(* IEC 61131-3 sources: daoli-st-library/DL_Process (part 69) *)

(* ---- FB_DL_PressFitStation.st ---- *)
(*==============================================================================
 * 组件名称 (Component)  : FB_DL_PressFitStation
 * 所属子库 (Sublibrary) : DL_Process
 * 当前版本 (Version)    : 1.0.0
 * 组件分类 (Category)   : 功能块（FUNCTION_BLOCK）· 工站模板 · 伺服精密压装
 * 兼容性 (Platform)     : CODESYS 3.5 / TwinCAT 3 / 汇川 InoProShop / Machine Expert；
 *                         仅依赖标准库（TON / R_TRIG / ABS / LIMIT / MAX / MIN），
 *                         位移与压力均为引脚注入的工程量，块内零硬件与零轴库细节
 * 功能描述 (Function)   : 伺服精密压装工站八态（待机 / 接近 / 压入 / 保压 / 回退 /
 *                         判定 / 完成 / 故障）；压入过程逐点做位移-压力包络窗口校验
 *                         （上下限按位移节点线性插值），提取接触点 / 屈服点 / 峰值点
 *                         / 终点四特征点，一个循环给出合格结论与 NG 原因位
 * 与既有件边界 (Scope)  : 轴级力矩限幅与到位判定属运动层力矩限幅件（只出「达限 /
 *                         到位」两个布尔）；本块做工站级工艺判定（包络 + 曲线特征 +
 *                         多原因归并 + 结果结构），分层不同、不可互替。通用步序基类
 *                         不套用：压装态与监控量强耦合，套基类会出现两套状态机并存
 * 状态机规模 (States)   : 八态最小子集（0 / 10 / 20 / 30 / 40 / 50 / 60 / 99），编号
 *                         留 10 间隔便于插态；不重复包装机十七态全集（那由包装机
 *                         状态机件承担），本块只做压装工序自身的可执行子集
 * 采样口径 (Sampling)   : 接近 / 压入 / 保压三段逐拍采样；包络校验只在压入与保压段
 *                         执行（接近段压力天然低于下限，一并判会误报）；斜率按相邻
 *                         两拍差分，位移增量小于保护阈值时沿用上一拍，杜绝除零
 * 屈服判据 (Yield note) : 取「斜率回落至峰值斜率的指定比例」，不以压力绝对过峰为前
 *                         提。现场屈服段多为斜率软化而非压力下降（铝壳 / 塑料件尤
 *                         甚），强求过峰则单调上升曲线永远判不出；过峰另有独立标志
 * 设计要点 (Key notes)  : ① 单拍三律：bDone 每拍预清零、eFinish 唯一置位、转出拍不
 *                           再置位；合格与不合格在 eEvaluate 一次锁存，同循环闭环
 *                         ② 包络表只读：注入表一律不改写，上下限对调在块内镜像纠正
 *                         ③ 二分定位：带防死锁计数的二分查找，节点上限 32，最多五轮
 *                         ④ 非有限值防御：位移或压力非有限时当拍拒绝采样并转故障
 *                         ⑤ 回退快照：进回退态首拍取终点特征，位置最多滞后一个扫描
 * 码位表 (Error codes)  :
 *   16#0005_01C0【信息级】包络表点数超上限已钳位为 32，不置故障位
 *   16#0005_01C1【信息级】包络上下限对调已在块内镜像修复，不置故障位
 *   16#0005_02C0【故障级】非法状态兜底
 *   16#0005_02C1【故障级】包络表非法（节点数小于 2、或位移非严格单调递增）
 *   16#0005_02C2【故障级】阶段超时（接近 / 压入 / 保压 三段共用该码）
 *   16#0005_02C3【故障级】采样非有限值（当拍拒绝更新并转故障）
 * NG 原因位 (NG bits)   : bit0 上包络越界｜bit1 下包络越界｜bit2 终点未达｜bit3 接触
 *                         未建立｜bit4 保压压降超限；按位或累计，一个循环可多位置位
 * R32 写入点次序审计 :
 *   nSampleCnt   : ① 启动拍清零（eIdle）→ ② 采样块自增（唯一自增点）
 *   uNgReason    : ① 启动拍清零 → ② 上包络越界 → ③ 下包络越界 → ④ 保压压降（eDwell
 *                  转出）→ ⑤ 终点未达（回退首拍）→ ⑥ 接触未建立（eEvaluate）→ ⑦ 复
 *                  位清；全部按位或置位，同拍按 ②③④⑤ 累加，结构上不可能互相覆盖
 *   _uErrorIdInt : ① 启动拍清零 → ② 包络表非法（启动校验）→ ③ 阶段超时（三态各一处，
 *                  同拍只命中一处）→ ④ 采样非有限 → ⑤ 非法状态（ELSE）→ ⑥ 复位清
 *   _eState      : 每拍只在 CASE 分支出口单点写入；CASE 之外仅两处（中止监视、使能撤
 *                  销），且均在 CASE 之前，次序固定
 * 验收向量 (Acceptance) :
 *   V1 包络插值：节点（0 毫米 上限 0 下限 0）、（10 毫米 上限 10 下限 2），实测位移
 *      5.0 毫米压力 5.5 千牛 → 插得上限 5.0 下限 1.0，上越界 0.5 千牛 → bit0 置位、
 *      最大偏差不小于 0.5 千牛（容差 1E-6）
 *   V2 接触点插值：采样（1.0 毫米, 0.02 千牛）、（1.2 毫米, 0.06 千牛），阈值 0.05
 *      千牛 → 接触位移 1.15 毫米（误差不超过 1E-4）
 *   V3 屈服点：斜率序列 20 / 18 / 9 千牛每毫米，比例 0.5（阈值 10）→ 斜率 9 出现那
 *      一拍锁存屈服点，锁存后不再更新
 *   V4 终点未达：目标 10.0 毫米，回退前最大位移 9.4 毫米 → bit2 置位、不合格、单拍脉冲
 *   V5 保压压降：保压起点 12.0 千牛、结束 8.0 千牛、判据 0.3 千牛 → 压降 4.0 千牛超限
 *      → bit4 置位
 *   V6 非法包络：节点数 1 → 码 02C1、故障锁存、不出完成脉冲
 * 开源溯源 (Origin)     : 参考 lisp 与 PLCopen 公开手册的「命令-监视-判定」三段分层与
 *                         工艺参数域命名组织，只借分类与参数域；状态机、插值、特征点
 *                         提取、码位与引脚契约为本库独立设计，clean-room 不构成衍生
 * 红线自检 (Redline)    : R1 零全局表与外部变量引用、零物理地址记号 ✓｜R2 零占位符 ✓
 *                         R3 纯 IEC 61131-3 加标准库 ✓｜R4 非有限值 / 除零 / 容差 /
 *                         判界 ✓｜R5 声明行中英双语同行注释 ✓｜R6 八成员逐一有 CASE
 *                         标签且含 ELSE 兜底 ✓｜R7 三沿两定时器 CASE 外无条件刷新 ✓
 * 修订历史 (Revision)   :
 *   2026-11-15  v1.0.0  首版入库（Round 11 · C 泳道 · 工站四件套之一）
 *============================================================================*)

(*------------------------------------------------------------------------------
 * 枚举: E_DL_PressFitState（归属 FB_DL_PressFitStation，同文件发布）
 *   八态：每个成员在下方主状态机中均有同名 CASE 标签，缺一即致命（R31）
 *-----------------------------------------------------------------------------*)
TYPE E_DL_PressFitState :
(
    eIdle      := 0,    // 待机：等启动沿，输出全复位 / Idle, awaiting start edge
    eApproach  := 10,   // 接近：等接触建立 / Approach, awaiting contact build-up
    ePress     := 20,   // 压入：包络校验与特征点逐拍提取 / Press, envelope and features per scan
    eDwell     := 30,   // 保压：保持压力并监视压降 / Dwell, hold and watch force decay
    eRetract   := 40,   // 回退：等回退到位或中止 / Retract, waiting for home or abort
    eEvaluate  := 50,   // 判定：归并 NG 原因并锁存结论 / Evaluate, merge NG reasons and latch
    eFinish    := 60,   // 完成：本拍出完成脉冲，下拍转待机 / Finish, done pulse this scan
    eFault     := 99    // 故障锁存：仅复位沿可退 / Fault latched, only a reset edge leaves
);
END_TYPE

(*------------------------------------------------------------------------------
 * 结构体: ST_DL_PressFitEnvelope（归属 FB_DL_PressFitStation）
 *   位移-压力包络表，由工艺组态注入；位移节点须严格单调递增
 *-----------------------------------------------------------------------------*)
TYPE ST_DL_PressFitEnvelope :
STRUCT
    nPoints   : INT;                        // 有效节点数 [个]，域 2~32 [Valid knot count]
    afPos     : ARRAY[1..32] OF REAL;       // 节点位移 [毫米]，严格单调递增 [Knot position, mm]
    afUpper   : ARRAY[1..32] OF REAL;       // 节点包络上限 [千牛] [Upper envelope limit, kN]
    afLower   : ARRAY[1..32] OF REAL;       // 节点包络下限 [千牛] [Lower envelope limit, kN]
END_STRUCT
END_TYPE

(*------------------------------------------------------------------------------
 * 结构体: ST_DL_PressFitResult（归属 FB_DL_PressFitStation）
 *   四特征点结果，未提取到时保持 0.0，对应 NG 原因位说明缺失原因
 *-----------------------------------------------------------------------------*)
TYPE ST_DL_PressFitResult :
STRUCT
    fContactPos   : REAL;                   // 接触点位移 [毫米] [Contact position, mm]
    fContactForce : REAL;                   // 接触点压力 [千牛] [Contact force, kN]
    fYieldPos     : REAL;                   // 屈服点位移 [毫米] [Yield position, mm]
    fYieldForce   : REAL;                   // 屈服点压力 [千牛] [Yield force, kN]
    fPeakPos      : REAL;                   // 峰值点位移 [毫米] [Peak position, mm]
    fPeakForce    : REAL;                   // 峰值点压力 [千牛] [Peak force, kN]
    fEndPos       : REAL;                   // 终点位移 [毫米] [End position, mm]
    fEndForce     : REAL;                   // 终点压力 [千牛] [End force, kN]
END_STRUCT
END_TYPE

(*------------------------------------------------------------------------------
 * 结构体: ST_DL_PressFitStat（归属 FB_DL_PressFitStation）
 *   跨周期统计，由调用方持有，本块只累加，掉电保持由上层负责
 *-----------------------------------------------------------------------------*)
TYPE ST_DL_PressFitStat :
STRUCT
    nCycleCount : UDINT;                    // 累计循环数 [次] [Cycle counter]
    nOkCount    : UDINT;                    // 累计合格数 [件] [Accepted counter]
    nNgCount    : UDINT;                    // 累计不合格数 [件] [Rejected counter]
END_STRUCT
END_TYPE

FUNCTION_BLOCK FB_DL_PressFitStation
VAR_INPUT
    bEnable            : BOOL;              // 使能，FALSE 回待机并复位输出 [Enable, FALSE resets to idle]
    bStart             : BOOL;              // 启动一个压装循环，上升沿受理 [Start one cycle on rising edge]
    bAbort             : BOOL;              // 中止并立即请求回退，上升沿受理 [Abort and retract on rising edge]
    bReset             : BOOL;              // 复位故障锁存，上升沿受理 [Reset latched fault on rising edge]
    fActPos            : REAL;              // 压头实际位移 [毫米]，量程 0.0~1000.0 [Ram position, mm]
    fActForce          : REAL;              // 压力传感器实测压力 [千牛]，量程 0.0~500.0 [Measured force, kN]
    fContactForceThr   : REAL := 0.05;      // 接触判定压力阈值 [千牛]，0 表示禁用接触点提取 [Contact threshold, kN]
    fYieldSlopeRatio   : REAL := 0.50;      // 屈服判据斜率比例 [-]，域 0.05~0.99 [Yield slope ratio]
    fPeakDropForce     : REAL := 0.30;      // 峰值后压降判定量 [千牛]，0 表示不判 [Force drop after peak, kN]
    fEndPosTarget      : REAL := 10.0;      // 终点位移目标 [毫米] [Target end position, mm]
    tStageTimeout      : TIME := T#5S;      // 单段动作超时 [毫秒]，0 表示不监控 [Per-stage timeout]
    tDwell             : TIME := T#500MS;   // 保压时间 [毫秒]，0 表示跳过保压 [Dwell time]
    fForceUpperLimit   : REAL := 180.0;     // 压力硬上限 [千牛]，达限立即转保压 [Hard force limit, kN]
END_VAR
VAR_OUTPUT
    eState             : E_DL_PressFitState; // 主状态机当前态 [-]，八态之一 [Current state]
    bBusy              : BOOL;              // 循环进行中，接近至回退为真 [Cycle in progress]
    bDone              : BOOL;              // 循环结束单拍脉冲 [-] [Single-scan done pulse]
    bOk                : BOOL;              // 判定合格，保持到下次启动 [Verdict OK held until next start]
    bNg                : BOOL;              // 判定不合格，保持到下次启动 [Verdict NG held until next start]
    bError             : BOOL;              // 故障级锁存，需复位清除 [Latched fault, cleared by reset]
    uErrorId           : UDINT;             // 事件码或故障码，0 表示无 [Event or fault code, 0 = none]
    uNgReason          : WORD;              // NG 原因位，bit0~bit4 见头注释 [NG reason bits, see header]
    stResult           : ST_DL_PressFitResult; // 曲线四特征点结果 [-] [Curve feature result]
    fEnvDevMax         : REAL;              // 全程包络最大偏差 [千牛]，趋势分析用 [Max envelope deviation, kN]
    nSampleCnt         : UDINT;             // 本循环有效采样点数 [点] [Valid sample count of this cycle]
END_VAR
VAR_IN_OUT
    stEnv              : ST_DL_PressFitEnvelope; // 包络表，组态注入，块内只读 [Envelope table, read-only here]
    stStat             : ST_DL_PressFitStat;     // 跨周期统计，调用方持有 [Persistent statistics held by caller]
END_VAR
VAR
    _eState            : E_DL_PressFitState := E_DL_PressFitState.eIdle; // 内部状态寄存器 [-]，唯一真值源 [Internal state register]
    _bInit             : BOOL := FALSE;     // 首扫标志，初值 FALSE，判据 NOT _bInit [First-scan flag, R19 pattern]
    _bFaultLatch       : BOOL;              // 故障级锁存，仅复位路径清 [Fault latch, reset path only]
    _uErrorIdInt       : UDINT;             // 故障级码寄存 [Fault-level code register]
    _uInfoCode         : UDINT;             // 本拍信息级码，每拍重算 [Transient info code]
    _bEnvValid         : BOOL;              // 包络表校验通过，启动拍重算 [Envelope validated at start]
    _nEnvPts           : INT;               // 生效包络节点数 [个]，域 2~32 [Effective knot count]
    _bContactFound     : BOOL;              // 接触点已提取 [Contact point captured]
    _bYieldFound       : BOOL;              // 屈服点已提取，只锁一次 [Yield point captured once]
    _bPeakPassed       : BOOL;              // 压力已回落过峰值 [Force passed its peak]
    _bHavePrev         : BOOL;              // 存在上一点采样 [Previous sample available]
    _bRetractSnapDone  : BOOL;              // 回退入口快照已完成 [Retract snapshot already taken]
    _fPrevPos          : REAL;              // 上一点位移 [毫米] [Previous position, mm]
    _fPrevForce        : REAL;              // 上一点压力 [千牛] [Previous force, kN]
    _fStartPos         : REAL;              // 循环起点位移 [毫米] [Cycle start position, mm]
    _fSlope            : REAL;              // 当前斜率 [千牛每毫米] [Current slope, kN/mm]
    _fSlopeMax         : REAL;              // 峰值斜率 [千牛每毫米] [Peak slope, kN/mm]
    _fPeakPos          : REAL;              // 峰值点位移 [毫米] [Peak position, mm]
    _fPeakForce        : REAL;              // 峰值点压力 [千牛] [Peak force, kN]
    _fDwellStartForce  : REAL;              // 保压起点压力 [千牛] [Dwell start force, kN]
    _fContactThrEff    : REAL;              // 生效接触阈值 [千牛] [Effective contact threshold, kN]
    _fYieldRatioEff    : REAL;              // 生效屈服比例 [-] [Effective yield ratio]
    _fPeakDropEff      : REAL;              // 生效压降判据 [千牛] [Effective drop criterion, kN]
    _fEndTgtEff        : REAL;              // 生效终点目标 [毫米] [Effective end target, mm]
    _fForceLimEff      : REAL;              // 生效压力硬上限 [千牛] [Effective force limit, kN]
    _tStageEff         : TIME;              // 生效单段超时 [毫秒] [Effective stage timeout]
    _tDwellEff         : TIME;              // 生效保压时间 [毫秒] [Effective dwell time]
    _fUp               : REAL;              // 插值包络上限 [千牛] [Interpolated upper bound, kN]
    _fLo               : REAL;              // 插值包络下限 [千牛] [Interpolated lower bound, kN]
    _fSpan             : REAL;              // 插值区间跨度 [毫米] [Interpolation span, mm]
    _fRatio            : REAL;              // 插值比例 [-] [Interpolation ratio]
    _fDelta            : REAL;              // 差分中间量 [千牛或毫米] [Difference term]
    afPosUse           : ARRAY[1..32] OF REAL;  // 位移节点镜像 [毫米] [Position knot mirror, mm]
    afUpperUse         : ARRAY[1..32] OF REAL;  // 包络上限镜像 [千牛] [Upper limit mirror, kN]
    afLowerUse         : ARRAY[1..32] OF REAL;  // 包络下限镜像 [千牛] [Lower limit mirror, kN]
    nI                 : INT;               // 通用循环索引 [索引] [Loop index]
    nGuard             : INT;               // 防死锁计数 [次] [Loop guard counter]
    nLo                : INT;               // 二分下界索引 [索引] [Binary search low index]
    nHi                : INT;               // 二分上界索引 [索引] [Binary search high index]
    nMid               : INT;               // 二分中点索引 [索引] [Binary search mid index]
    bSampleFinite      : BOOL;              // 采样值有限，当拍可采 [Sample finite verdict]
    _bStageChg         : BOOL;              // 本拍发生过阶段迁移，用于断开单段计时一拍 [Stage changed this scan]
    _eStagePrev        : E_DL_PressFitState := E_DL_PressFitState.eIdle; // 上拍状态，迁移判据用 [Previous state of last scan]
    bStageTmoIn        : BOOL;              // 单段超时输入条件，先算后调 [Stage timer input]
    bDwellTmoIn        : BOOL;              // 保压计时输入条件，先算后调 [Dwell timer input]
    fbTrigStart        : R_TRIG;            // 启动沿检测 [Start edge detector]
    fbTrigAbort        : R_TRIG;            // 中止沿检测 [Abort edge detector]
    fbTrigReset        : R_TRIG;            // 复位沿检测 [Reset edge detector]
    fbTmoStage         : TON;               // 单段超时定时器 [Stage timeout timer]
    fbTmoDwell         : TON;               // 保压计时定时器 [Dwell timer]
END_VAR
VAR CONSTANT
    DL_FLOAT_EPS       : REAL := 1.0E-6;    // 浮点判等容差 [-] [Float comparison epsilon]
    DL_SLOPE_MIN_DELTA : REAL := 1.0E-4;    // 斜率计算最小位移增量 [毫米] [Min delta for slope, mm]
    DL_ENV_MAX_POINTS  : INT  := 32;        // 包络表节点数上限 [个] [Max envelope knots]
    DL_ENV_MIN_POINTS  : INT  := 2;         // 包络表节点数下限 [个] [Min envelope knots]
    DL_MAX_LOOP        : INT  := 64;        // 循环防死锁上限 [次] [Loop guard limit]
    DL_MAX_CYCLES      : UDINT := 16#FFFF_FFFE; // 统计计数饱和上限 [次] [Counter saturation limit]
    DL_RATIO_MIN       : REAL := 0.05;      // 屈服比例域下限 [-] [Yield ratio lower bound]
    DL_RATIO_MAX       : REAL := 0.99;      // 屈服比例域上限 [-] [Yield ratio upper bound]
    DL_FORCE_MAX       : REAL := 500.0;     // 压力输入域上限 [千牛] [Force domain upper bound, kN]
    DL_POS_MAX         : REAL := 1000.0;    // 位移输入域上限 [毫米] [Position domain upper bound, mm]
    DL_REAL_MAX        : REAL := 3.4E38;    // 单精度有限值判据幅值 [-] [Finite magnitude bound]
    DL_TMO_MAX         : TIME := T#180S;    // 超时参数域上限 [毫秒] [Timeout upper bound]
    DL_NG_ENV_HIGH     : WORD := 16#0001;   // NG 原因位 bit0 上包络越界 [NG bit0, upper envelope]
    DL_NG_ENV_LOW      : WORD := 16#0002;   // NG 原因位 bit1 下包络越界 [NG bit1, lower envelope]
    DL_NG_END_POS      : WORD := 16#0004;   // NG 原因位 bit2 终点未达 [NG bit2, end not reached]
    DL_NG_NO_CONTACT   : WORD := 16#0008;   // NG 原因位 bit3 接触未建立 [NG bit3, contact missing]
    DL_NG_DWELL_DROP   : WORD := 16#0010;   // NG 原因位 bit4 保压压降超限 [NG bit4, dwell decay]
    DL_INFO_PTS_CLAMP  : UDINT := 16#0005_01C0; // 01C0 包络点数越界已钳位【信息级】 [Info, knots clamped]
    DL_INFO_LIM_SWAP   : UDINT := 16#0005_01C1; // 01C1 上下限对调已修复【信息级】 [Info, limits swapped]
    DL_ERR_STATE       : UDINT := 16#0005_02C0; // 02C0 非法状态兜底【故障级】 [Fault, illegal state]
    DL_ERR_ENV         : UDINT := 16#0005_02C1; // 02C1 包络表非法【故障级】 [Fault, invalid envelope]
    DL_ERR_STAGE_TMO   : UDINT := 16#0005_02C2; // 02C2 阶段超时【故障级】 [Fault, stage timeout]
    DL_ERR_SAMPLE      : UDINT := 16#0005_02C3; // 02C3 采样非有限值【故障级】 [Fault, non-finite sample]
END_VAR
// ==== 段 1｜单拍输出预清零（R24/R25 律①：置位前先清零，任何早退路径输出确定） / Single-scan output pre-clear, mandatory before any set point
bDone      := FALSE;                        // 完成脉冲每拍先清零 [Done pulse pre-cleared]
_uInfoCode := 16#0000_0000;                 // 信息级码每拍重算 [Info code recomputed each scan]
// ==== 段 2｜工艺参数钳位（先钳位再进逻辑，杜绝分支内出现裸数值） / Parameter clamping before any logical use, no magic numbers in logic
_fContactThrEff := LIMIT(0.0, fContactForceThr, DL_FORCE_MAX);   // 接触阈值钳位 [千牛] [Contact threshold clamped]
_fYieldRatioEff := LIMIT(DL_RATIO_MIN, fYieldSlopeRatio, DL_RATIO_MAX); // 屈服比例钳位 [-] [Yield ratio clamped]
_fPeakDropEff   := LIMIT(0.0, fPeakDropForce, DL_FORCE_MAX);     // 压降判据钳位 [千牛] [Drop criterion clamped]
_fEndTgtEff     := LIMIT(0.0, fEndPosTarget, DL_POS_MAX);        // 终点目标钳位 [毫米] [End target clamped]
_fForceLimEff   := LIMIT(DL_FLOAT_EPS, fForceUpperLimit, DL_FORCE_MAX); // 硬上限钳位 [千牛] [Force limit clamped]
_tStageEff := tStageTimeout;                // 单段超时先取引脚值 [Stage timeout from pin]
IF _tStageEff > DL_TMO_MAX THEN
    _tStageEff := DL_TMO_MAX;               // 超上限钳位 [Clamped to upper bound]
ELSIF _tStageEff < T#0S THEN
    _tStageEff := T#0S;                     // 负值归零 [Negative clamped to zero]
END_IF
_tDwellEff := tDwell;                       // 保压时间先取引脚值 [Dwell time from pin]
IF _tDwellEff > DL_TMO_MAX THEN
    _tDwellEff := DL_TMO_MAX;               // 超上限钳位 [Clamped to upper bound]
ELSIF _tDwellEff < T#0S THEN
    _tDwellEff := T#0S;                     // 负值归零 [Negative clamped to zero]
END_IF
// ==== 段 3｜沿与定时器无条件刷新（R7 红线：严禁置于 IF / CASE 分支内） / Unconditional per-cycle refresh of edges and timers, outside any branch
fbTrigStart(CLK := bStart);                 // 启动沿 [Start edge]
fbTrigAbort(CLK := bAbort);                 // 中止沿 [Abort edge]
fbTrigReset(CLK := bReset);                 // 复位沿 [Reset edge]
IF ((_eState = E_DL_PressFitState.eApproach)
 OR (_eState = E_DL_PressFitState.ePress)
 OR (_eState = E_DL_PressFitState.eDwell)) AND (NOT _bStageChg) THEN
    bStageTmoIn := TRUE;                    // 动作段计时，迁移后的第一拍断输入以清零 [Timed, broken one scan after a transition]
ELSE
    bStageTmoIn := FALSE;                   // 非动作段不计时 [Timer disabled outside motion]
END_IF
fbTmoStage(IN := bStageTmoIn, PT := _tStageEff);
IF _eState = E_DL_PressFitState.eDwell THEN
    bDwellTmoIn := TRUE;                    // 仅保压段计时 [Only during dwell]
ELSE
    bDwellTmoIn := FALSE;                   // 其余段清零 [Cleared otherwise]
END_IF
fbTmoDwell(IN := bDwellTmoIn, PT := _tDwellEff);
// ==== 段 4｜首扫初始化（R19 唯一合法范式：初值 FALSE，判据 NOT，同步后置 TRUE） / First-scan initialisation with the canonical R19 pattern
IF NOT _bInit THEN
    _eState           := E_DL_PressFitState.eIdle;  // 状态回待机 [State to idle]
    _bFaultLatch      := FALSE;             // 故障锁存清零 [Fault latch cleared]
    _uErrorIdInt      := 16#0000_0000;      // 故障码清零 [Fault code cleared]
    _bEnvValid        := FALSE;             // 包络未校验 [Envelope not validated yet]
    _bStageChg        := FALSE;             // 阶段迁移标志清零 [Stage change flag cleared]
    _eStagePrev       := E_DL_PressFitState.eIdle;  // 上拍状态同步 [Previous state synced]
    _nEnvPts          := 0;                 // 节点数清零 [Knot count cleared]
    _bContactFound    := FALSE;  _bYieldFound   := FALSE;   // 接触点与屈服点未提取 [Contact and yield not captured]
    _bPeakPassed      := FALSE;  _bHavePrev     := FALSE;   // 过峰标志与采样链清零 [Peak flag and sampling chain cleared]
    _bRetractSnapDone := FALSE;             // 回退快照未做 [Retract snapshot pending]
    _fPrevPos         := 0.0;    _fPrevForce    := 0.0;     // 上一点位移与压力清零 [Previous sample cleared]
    _fStartPos        := 0.0;    _fDwellStartForce := 0.0;  // 起点与保压起点压力清零 [Start points cleared]
    _fSlope           := 0.0;    _fSlopeMax     := 0.0;     // 斜率与峰值斜率清零 [Slope and peak slope cleared]
    _fPeakPos         := 0.0;    _fPeakForce    := 0.0;     // 峰值点清零 [Peak point cleared]
    fEnvDevMax        := 0.0;    _fUp           := 0.0;     // 最大偏差与插值上限清零 [Deviation and upper bound cleared]
    _fLo              := 0.0;                               // 插值下限清零 [Lower bound cleared]
    bOk               := FALSE;  bNg            := FALSE;   // 合格与不合格结论清零 [Verdicts cleared]
    bBusy             := FALSE;  bError         := FALSE;   // 忙与故障标志清零 [Busy and error cleared]
    uErrorId          := 16#0000_0000;  uNgReason := 16#0000;  // 事件码与原因位清零 [Error id and NG bits cleared]
    nSampleCnt        := 0;                 // 采样计数清零 [Sample counter cleared]
    stResult.fContactPos   := 0.0;  stResult.fContactForce := 0.0;  // 接触点清零 [Contact point cleared]
    stResult.fYieldPos     := 0.0;  stResult.fYieldForce   := 0.0;  // 屈服点清零 [Yield point cleared]
    stResult.fPeakPos      := 0.0;  stResult.fPeakForce    := 0.0;  // 峰值点清零 [Peak point cleared]
    stResult.fEndPos       := 0.0;  stResult.fEndForce     := 0.0;  // 终点清零 [End point cleared]
    FOR nI := 1 TO DL_ENV_MAX_POINTS DO
        afPosUse[nI]   := 0.0;              // 位移镜像清零 [Position mirror cleared]
        afUpperUse[nI] := 0.0;              // 上限镜像清零 [Upper mirror cleared]
        afLowerUse[nI] := 0.0;              // 下限镜像清零 [Lower mirror cleared]
    END_FOR
    _bInit := TRUE;                         // 首扫只做一次 [Runs exactly once]
END_IF
// ==== 段 5｜启动拍包络表校验（只读校验，上下限对调在镜像里纠正，绝不改写组态） / Envelope validation at start; swaps are repaired in the mirror only
IF fbTrigStart.Q AND (_eState = E_DL_PressFitState.eIdle)
AND bEnable AND (NOT _bFaultLatch) THEN
    _bEnvValid := TRUE;                     // 先假定合法，再逐条反证 [Assume valid, then disprove]
    _nEnvPts   := stEnv.nPoints;            // 取组态节点数 [Knot count from configuration]
    IF _nEnvPts > DL_ENV_MAX_POINTS THEN
        _nEnvPts   := DL_ENV_MAX_POINTS;    // 超上限钳到 32 [Clamped to 32]
        _uInfoCode := DL_INFO_PTS_CLAMP;    // 01C0 点数越界已钳位【信息级】 [Info, knots clamped]
    END_IF
    IF _nEnvPts < DL_ENV_MIN_POINTS THEN
        _bEnvValid := FALSE;                // 少于两点无法插值 [Less than two knots is unusable]
    END_IF
    IF _bEnvValid THEN
        FOR nI := 1 TO _nEnvPts DO
            afPosUse[nI] := stEnv.afPos[nI];    // 位移镜像复制 [Copy position knot]
            IF stEnv.afUpper[nI] < stEnv.afLower[nI] THEN
                afUpperUse[nI] := stEnv.afLower[nI];   // 上限取原下限 [Upper takes old lower]
                afLowerUse[nI] := stEnv.afUpper[nI];   // 下限取原上限 [Lower takes old upper]
                _uInfoCode     := DL_INFO_LIM_SWAP;    // 01C1 上下限对调已修复【信息级】 [Info, limits swapped]
            ELSE
                afUpperUse[nI] := stEnv.afUpper[nI];  afLowerUse[nI] := stEnv.afLower[nI];  // 正常复制上下限 [Copy limits as-is]
            END_IF
        END_FOR
        FOR nI := 1 TO (_nEnvPts - 1) DO
            IF afPosUse[nI + 1] <= afPosUse[nI] THEN
                _bEnvValid := FALSE;        // 位移非严格单调，二分不可用 [Non-monotonic, binary search unsafe]
            END_IF
        END_FOR
    END_IF
    IF NOT _bEnvValid THEN
        _bFaultLatch := TRUE;               // 故障锁存 [Fault latched]
        _uErrorIdInt := DL_ERR_ENV;         // 02C1 包络表非法【故障级】 [Fault, invalid envelope]
        _eState      := E_DL_PressFitState.eFault;
    END_IF
END_IF
// ==== 段 6｜采样有限性防御与中止监视（全局，优先于状态机） / Sample finiteness defense and abort monitor, ahead of the state machine
bSampleFinite := (fActPos >= (-DL_REAL_MAX)) AND (fActPos <= DL_REAL_MAX)
             AND (fActForce >= (-DL_REAL_MAX)) AND (fActForce <= DL_REAL_MAX);
IF bEnable AND (NOT _bFaultLatch)
AND (_eState <> E_DL_PressFitState.eIdle)
AND (_eState <> E_DL_PressFitState.eFault)
AND (NOT bSampleFinite) THEN
    _bFaultLatch := TRUE;                   // 非有限值属故障级，立即锁存 [Non-finite is a fault]
    _uErrorIdInt := DL_ERR_SAMPLE;          // 02C3 采样非有限值【故障级】 [Fault, non-finite sample]
    _eState      := E_DL_PressFitState.eFault;
END_IF

IF bEnable AND (NOT _bFaultLatch) AND fbTrigAbort.Q
AND ((_eState = E_DL_PressFitState.eApproach)
  OR (_eState = E_DL_PressFitState.ePress)
  OR (_eState = E_DL_PressFitState.eDwell)) THEN
    _bHavePrev := FALSE;                    // 中止后重新起算差分 [Difference restarts after abort]
    _eState    := E_DL_PressFitState.eRetract;
END_IF
// ==== 段 7｜使能撤销（FALSE 立即回待机并撤全部动作出口，保留故障锁存） / Disable path returns to idle immediately, fault latch is preserved
IF NOT bEnable THEN
    _eState      := E_DL_PressFitState.eIdle;
    _bHavePrev   := FALSE;                  // 采样链断，防跨循环沿用 [Sampling chain broken]
    bBusy        := FALSE;                  // 忙标志撤 [Busy withdrawn]
END_IF
// ==== 段 8｜采样与特征点提取（接近 / 压入 / 保压三段逐拍执行） / Sampling and feature extraction, one sample per scan in three stages
IF bEnable AND (NOT _bFaultLatch) AND bSampleFinite
AND ((_eState = E_DL_PressFitState.eApproach)
  OR (_eState = E_DL_PressFitState.ePress)
  OR (_eState = E_DL_PressFitState.eDwell)) THEN

    IF _bHavePrev THEN
        // ---- 斜率：相邻两拍差分，位移增量过小时沿用上一拍，杜绝除零
        _fDelta := fActPos - _fPrevPos;
        IF ABS(_fDelta) >= DL_SLOPE_MIN_DELTA THEN
            _fSlope := (fActForce - _fPrevForce) / _fDelta;   // 斜率 [千牛每毫米] [Slope, kN/mm]
        END_IF
        IF _fSlope > _fSlopeMax THEN
            _fSlopeMax := _fSlope;          // 跟踪峰值斜率 [Track peak slope]
        END_IF
        // ---- 接触点：首个越过阈值的采样，用相邻两采样线性插值求精确位移
        IF (NOT _bContactFound) AND (_fContactThrEff > DL_FLOAT_EPS)
        AND (fActForce >= _fContactThrEff) THEN
            _fDelta := fActForce - _fPrevForce;
            IF ABS(_fDelta) > DL_FLOAT_EPS THEN
                stResult.fContactPos := _fPrevPos
                    + (fActPos - _fPrevPos) * (_fContactThrEff - _fPrevForce) / _fDelta;
            ELSE
                stResult.fContactPos := fActPos;   // 压力已稳定在阈值上，退化为当前点 [Degenerate to current point]
            END_IF
            stResult.fContactForce := fActForce;   // 接触点压力 [Contact force, kN]
            _bContactFound         := TRUE;        // 只锁一次 [Latched once]
        END_IF
    END_IF

    // ---- 峰值点：全程最大压力及其位移，逐拍刷新
    IF fActForce > _fPeakForce THEN
        _fPeakForce        := fActForce;    // 峰值压力 [千牛] [Peak force, kN]
        _fPeakPos          := fActPos;      // 峰值位移 [毫米] [Peak position, mm]
        stResult.fPeakForce := _fPeakForce;
        stResult.fPeakPos   := _fPeakPos;
    END_IF
    IF fActForce < (_fPeakForce - DL_FLOAT_EPS) THEN
        _bPeakPassed := TRUE;               // 已回落过峰值，趋势用 [Force has passed its peak]
    END_IF

    // ---- 屈服点：斜率回落至峰值斜率指定比例，首次成立即锁存
    IF (NOT _bYieldFound) AND _bContactFound AND (_fSlopeMax > DL_FLOAT_EPS) THEN
        IF _fSlope < (_fSlopeMax * _fYieldRatioEff) THEN
            stResult.fYieldPos   := fActPos;    // 屈服位移 [毫米] [Yield position, mm]
            stResult.fYieldForce := fActForce;  // 屈服压力 [千牛] [Yield force, kN]
            _bYieldFound         := TRUE;       // 只锁一次 [Latched once]
        END_IF
    END_IF

    nSampleCnt := nSampleCnt + 1;           // 有效采样计数 [Valid sample counter]
    _fPrevPos  := fActPos;                  // 上一点位移刷新 [Previous position refreshed]
    _fPrevForce := fActForce;               // 上一点压力刷新 [Previous force refreshed]
    _bHavePrev := TRUE;                     // 已有上一点 [Previous sample available]

    // ---- 包络窗口校验：仅压入与保压段，接近段压力天然低于下限故不判
    IF (_eState = E_DL_PressFitState.ePress) OR (_eState = E_DL_PressFitState.eDwell) THEN
        nLo    := 1;
        nHi    := _nEnvPts;
        nGuard := 0;
        WHILE ((nHi - nLo) > 1) AND (nGuard < DL_MAX_LOOP) DO
            nGuard := nGuard + 1;           // 防死锁计数 [Guard incremented]
            nMid   := (nLo + nHi) / 2;      // 整数中点 [Integer midpoint]
            IF fActPos >= afPosUse[nMid] THEN
                nLo := nMid;                // 落在右半区 [Right half]
            ELSE
                nHi := nMid;                // 落在左半区 [Left half]
            END_IF
        END_WHILE
        _fSpan := afPosUse[nHi] - afPosUse[nLo];
        IF ABS(_fSpan) > DL_SLOPE_MIN_DELTA THEN
            _fRatio := (fActPos - afPosUse[nLo]) / _fSpan;         // 区间内比例 [-] [Ratio in interval]
            _fRatio := LIMIT(0.0, _fRatio, 1.0);                   // 区间外钳位 [Clamped to 0..1]
            _fUp := afUpperUse[nLo] + _fRatio * (afUpperUse[nHi] - afUpperUse[nLo]); // 插值上限 [Interpolated upper]
            _fLo := afLowerUse[nLo] + _fRatio * (afLowerUse[nHi] - afLowerUse[nLo]); // 插值下限 [Interpolated lower]
        ELSE
            _fUp := afUpperUse[nLo];        // 退化区间取左节点上限 [Degenerate, take left knot]
            _fLo := afLowerUse[nLo];        // 退化区间取左节点下限 [Degenerate, take left knot]
        END_IF
        IF fActForce > (_fUp + DL_FLOAT_EPS) THEN
            uNgReason := uNgReason OR DL_NG_ENV_HIGH;              // bit0 上包络越界 [Upper envelope violated]
            IF (fActForce - _fUp) > fEnvDevMax THEN
                fEnvDevMax := fActForce - _fUp;                    // 累计最大偏差 [Track max deviation]
            END_IF
        END_IF
        IF fActForce < (_fLo - DL_FLOAT_EPS) THEN
            uNgReason := uNgReason OR DL_NG_ENV_LOW;               // bit1 下包络越界 [Lower envelope violated]
            IF (_fLo - fActForce) > fEnvDevMax THEN
                fEnvDevMax := _fLo - fActForce;                    // 累计最大偏差 [Track max deviation]
            END_IF
        END_IF
    END_IF
END_IF
// ==== 段 9｜主状态机（ENUM 加 CASE 加 ELSE 兜底，八成员逐一有标签） / Main state machine, every enum member has its own label
CASE _eState OF
    E_DL_PressFitState.eIdle: // 待机：等启动沿，启动拍清循环量
        IF fbTrigStart.Q AND bEnable AND (NOT _bFaultLatch) AND _bEnvValid THEN
            uNgReason    := 16#0000;  fEnvDevMax := 0.0;  nSampleCnt := 0;   // 原因位、最大偏差、采样计数清零 [Bits, deviation, count cleared]
            _bContactFound := FALSE;  _bYieldFound := FALSE;  _bPeakPassed := FALSE;  // 特征点与过峰标志复位 [Feature flags reset]
            _bHavePrev := FALSE;      _fSlope := 0.0;   _fSlopeMax := 0.0;         // 采样链、斜率、峰值斜率复位 [Chain and slope reset]
            _fPeakPos := 0.0;         _fPeakForce := 0.0;                          // 峰值点复位 [Peak reset]
            _fStartPos := fActPos;    _bRetractSnapDone := FALSE;                  // 记循环起点并复位回退快照 [Start point and snapshot reset]
            _uErrorIdInt := 16#0000_0000;  bOk := FALSE;  bNg := FALSE;            // 故障码与结论复位（启动前必无故障）[Code and verdicts reset]
            stResult.fContactPos := 0.0;  stResult.fContactForce := 0.0;           // 接触点复位 [Contact reset]
            stResult.fYieldPos   := 0.0;  stResult.fYieldForce   := 0.0;           // 屈服点复位 [Yield reset]
            stResult.fPeakPos    := 0.0;  stResult.fPeakForce    := 0.0;           // 峰值点复位 [Peak reset]
            stResult.fEndPos     := 0.0;  stResult.fEndForce     := 0.0;           // 终点复位 [End reset]
            _eState := E_DL_PressFitState.eApproach;
        END_IF
    E_DL_PressFitState.eApproach: // 接近：接触建立即转压入，阈值禁用时直通
        IF (_fContactThrEff <= DL_FLOAT_EPS) OR _bContactFound THEN
            _eState := E_DL_PressFitState.ePress;
        ELSIF fbTmoStage.Q THEN
            _bFaultLatch := TRUE;           // 阶段超时锁存 [Stage timeout latched]
            _uErrorIdInt := DL_ERR_STAGE_TMO;  // 02C2 阶段超时【故障级】 [Fault, stage timeout]
            _eState      := E_DL_PressFitState.eFault;
        END_IF
    E_DL_PressFitState.ePress: // 压入：到达终点目标或压力硬上限即转保压
        IF (fActPos >= (_fEndTgtEff - DL_FLOAT_EPS)) OR (fActForce >= _fForceLimEff) THEN
            _fDwellStartForce := fActForce; // 保压起点压力快照 [Dwell start force snapshot]
            _eState           := E_DL_PressFitState.eDwell;
        ELSIF fbTmoStage.Q THEN
            _bFaultLatch := TRUE;           // 阶段超时锁存 [Stage timeout latched]
            _uErrorIdInt := DL_ERR_STAGE_TMO;  // 02C2 阶段超时【故障级】 [Fault, stage timeout]
            _eState      := E_DL_PressFitState.eFault;
        END_IF
    E_DL_PressFitState.eDwell: // 保压：计时到即判压降并转回退，零时长直通
        IF (_tDwellEff <= T#0S) OR fbTmoDwell.Q THEN
            IF (_fPeakDropEff > DL_FLOAT_EPS)
            AND ((_fDwellStartForce - fActForce) > _fPeakDropEff) THEN
                uNgReason := uNgReason OR DL_NG_DWELL_DROP;  // bit4 保压压降超限 [Dwell decay violated]
            END_IF
            _bHavePrev := FALSE;            // 回退段不再算斜率 [Slope tracking stops]
            _eState    := E_DL_PressFitState.eRetract;
        ELSIF fbTmoStage.Q THEN
            _bFaultLatch := TRUE;           // 阶段超时锁存 [Stage timeout latched]
            _uErrorIdInt := DL_ERR_STAGE_TMO;  // 02C2 阶段超时【故障级】 [Fault, stage timeout]
            _eState      := E_DL_PressFitState.eFault;
        END_IF
    E_DL_PressFitState.eRetract: // 回退：首拍取终点特征，到位或中止即转判定
        IF NOT _bRetractSnapDone THEN
            stResult.fEndPos   := fActPos;  // 终点位移 [毫米] [End position, mm]
            stResult.fEndForce := fActForce; // 终点压力 [千牛] [End force, kN]
            IF fActPos < (_fEndTgtEff - DL_FLOAT_EPS) THEN
                uNgReason := uNgReason OR DL_NG_END_POS;  // bit2 终点未达 [End position not reached]
            END_IF
            _bRetractSnapDone := TRUE;      // 快照只做一次 [Snapshot taken once]
        END_IF
        IF fbTrigAbort.Q OR (fActPos <= (_fStartPos + DL_FLOAT_EPS)) THEN
            _eState := E_DL_PressFitState.eEvaluate;
        END_IF
    E_DL_PressFitState.eEvaluate: // 判定：归并原因并锁存结论，当拍转完成
        IF (_fContactThrEff > DL_FLOAT_EPS) AND (NOT _bContactFound) THEN
            uNgReason := uNgReason OR DL_NG_NO_CONTACT;  // bit3 接触未建立 [Contact never built up]
        END_IF
        bNg      := (uNgReason <> 16#0000); // 任一原因位即不合格 [Any reason bit means NG]
        bOk      := NOT bNg;                // 与不合格严格互斥 [Mutually exclusive with NG]
        _eState  := E_DL_PressFitState.eFinish;
    E_DL_PressFitState.eFinish: // 完成：本拍出完成脉冲并结算统计，下拍转待机
        bDone := TRUE;                      // 完成单拍，本拍唯一置位点 [Sole set point of the pulse]
        IF bNg THEN
            IF stStat.nNgCount < DL_MAX_CYCLES THEN
                stStat.nNgCount := stStat.nNgCount + 1;   // 不合格计数饱和累加 [NG counter, saturated]
            END_IF
        ELSE
            IF stStat.nOkCount < DL_MAX_CYCLES THEN
                stStat.nOkCount := stStat.nOkCount + 1;   // 合格计数饱和累加 [OK counter, saturated]
            END_IF
        END_IF
        IF stStat.nCycleCount < DL_MAX_CYCLES THEN
            stStat.nCycleCount := stStat.nCycleCount + 1; // 循环计数饱和累加 [Cycle counter, saturated]
        END_IF
        _bHavePrev := FALSE;                // 采样链断开，防跨循环 [Sampling chain broken]
        _eState    := E_DL_PressFitState.eIdle;
    E_DL_PressFitState.eFault: // 故障：等复位沿，复位后清码回待机
        IF fbTrigReset.Q THEN
            _bFaultLatch      := FALSE;     // 锁存解除 [Latch released]
            _uErrorIdInt      := 16#0000_0000; // 故障码清零 [Fault code cleared]
            uNgReason         := 16#0000;   // 原因位清零 [NG bits cleared]
            _bRetractSnapDone := FALSE;     // 快照标志复位 [Snapshot flag reset]
            _bHavePrev        := FALSE;     // 差分复位 [Difference reset]
            _eState           := E_DL_PressFitState.eIdle;
        END_IF

    ELSE // 非法枚举值兜底：回安全态并锁故障
        _bFaultLatch := TRUE;               // 兜底锁存 [Fallback latch]
        _uErrorIdInt := DL_ERR_STATE;       // 02C0 非法状态兜底【故障级】 [Fault, illegal state]
        _eState      := E_DL_PressFitState.eFault;
END_CASE
// ==== 段 10｜阶段迁移寄存器更新（单段超时的清零依据，与状态写入点分离） / Stage change register, drives the per-stage timer reset
_bStageChg  := (_eState <> _eStagePrev);     // 本拍是否发生迁移 [Transition happened this scan]
_eStagePrev := _eState;                      // 迁移寄存器同步 [Previous state synced]

// ==== 段 11｜出口派生（每拍重写，bError 只反映故障级，信息级码只进 uErrorId） / Outlets rewritten every scan, info codes never raise bError
eState := _eState;                          // 状态镜像 [State mirror]
bBusy  := (_eState = E_DL_PressFitState.eApproach)
       OR (_eState = E_DL_PressFitState.ePress)
       OR (_eState = E_DL_PressFitState.eDwell)
       OR (_eState = E_DL_PressFitState.eRetract);   // 执行中派生 [Busy derived]

bError := _bFaultLatch;                     // 故障级派生式（R21）[Fault-level derived form]
IF _bFaultLatch THEN
    uErrorId := _uErrorIdInt;               // 故障级码优先透出 [Fault code wins]
ELSE
    uErrorId := _uInfoCode;                 // 无故障时透出信息级码 [Info code otherwise]
END_IF
END_FUNCTION_BLOCK

(* ---- FB_DL_PressForceCurveExec.st ---- *)
(*==============================================================================
 * 组件名称 (Component)  : FB_DL_PressForceCurveExec
 * 所属子库 (Sublibrary) : DL_Process ｜ 版本 (Version) : 1.0.0 ｜ 2026-11-24
 * 兼容性   (Platform)   : CODESYS 3.5+ / TwinCAT 3 / 汇川 InoProShop / 施耐德 Machine Expert
 *                         仅依赖 IEC 61131-3 标准库（TON / R_TRIG / ABS / MIN / MAX / LIMIT），零厂商私有库
 * 功能描述 (Function)   : 压机多段力曲线执行：按 4 段配方（目标力 aSegForce / 升力速率 aSegRate /
 *                         保压时长 aSegHold）逐段执行，eRamp 以「速率 × dt」斜坡逼近目标力，
 *                         到力判据 = 指令已饱和到目标（|cmd − target| ≤ EPS）**且** 实际力反馈落进
 *                         容差带（容差 = max(0.5% × |目标力|, 0.1 kN)）→ eHold 保压 aSegHold[i]；
 *                         末段保压完成 → eRelease 按末段速率把力指令斜坡降到 0 → eDone 发 bCurveDone。
 *                         **dt 口径**：定周期采样节拍 tonDt（PT = 100ms 常数）生成步长
 *                         _fDtSec := TIME_TO_LREAL(DL_PFC_DT)，入口做 dt > EPS 闸（R4 防 dt ≤ 0）；
 *                         保压计时用 DINT 毫秒累加（_diHoldMs，每采样拍 +100ms），避免 TIME 加法跨型。
 *                         **bStart = FALSE 语义（R191 二选一，本件选「降级为安全值 + 置标志」）**：
 *                         力指令按段速率退回 0 并进 eIdle（压机力指令不得冻结保持）。
 * 接口     (Interface)  : 输入 bEnable / bStart / bReset（上升沿）/ aSegForce[1..4] / aSegRate[1..4] /
 *                         aSegHold[1..4] / nSegCnt / fForceFb / tSegTimeout；
 *                         输出 fForceCmd / nSegAct / tHoldElapsed / bCurveDone / eState（E_DL_PfcPhase）/
 *                         eCause（E_DL_PfcCause）/ bError / bValid / nSegCompleted。
 * 状态迁移表 (State Transition Table)：
 *   ① eIdle → eRamp：bEnable 且 bStart 且组态闸通过且无锁存；拍 N 进入 / 本拍行为：
 *      fForceCmd=0、nSegAct=1、nSegCompleted=0、_diHoldMs=0 / 拍 N+1 转出至 eRamp。
 *   ② eRamp → eHold：到力判据成立（指令饱和 + 反馈落带）；拍 N 进入 / 本拍行为：
 *      _diHoldMs 清零、fForceCmd 精确取目标 / 拍 N+1 转出至 eHold。
 *   ③ eHold → eRamp：_diHoldMs ≥ aSegHold[i] 且 i < nSegCnt；本拍行为：nSegAct+1、
 *      nSegCompleted+1、_diHoldMs 清零、信息级 eSegDone / 拍 N+1 转出（下一段）。
 *   ④ eHold → eRelease：_diHoldMs ≥ aSegHold[nSegCnt]（末段完成）；本拍行为：nSegCompleted+1、
 *      信息级 eCurveDoneCode / 拍 N+1 转出至 eRelease。
 *   ⑤ eRelease → eDone：|fForceCmd| ≤ EPS（已退到 0）；本拍行为：fForceCmd 精确置 0 /
 *      拍 N+1 转出至 eDone。
 *   ⑥ eDone → eIdle：(NOT bStart) OR bReset 上升沿（两条出口 R98）；本拍行为：bCurveDone 落 FALSE、
 *      力指令与段号清零 / 拍 N+1 转出至 eIdle。
 *   ⑦ eRamp → eFault：tonSeg.Q（单段超时未到力）锁存 eForceNotReached；本拍行为：fForceCmd 保持
 *      当前值直至段尾迁移闸（R21）后再全撤 / 拍 N+1 转出至 eFault。
 *   ⑧ 任一相 → eFault：组态闸失败（段数越域 / 速率 ≤ 0 / 目标力 < 0 / 保压越域 / 超时越域 /
 *      fForceFb 非有限），锁存首因。
 *   ⑨ eFault → eIdle：bReset 上升沿（R_TRIG 判 .Q）且 bEnable = FALSE（R19 穷举出口）；
 *      本拍行为：清锁存与成因、fForceCmd=0 / 拍 N+1 转出至 eIdle。
 *   ⑩ ELSE（非法枚举值）→ eFault，成因 eIllegalState（R6 兜底）。
 * 边界     (Boundary)   : ① tonDt / tonSeg / R_TRIG 全在 CASE 外无条件调用（R7）；两者 IN 均含
 *                            NOT .Q 自复位项（R188）；tonSeg 另含「(NOT _bSegReset)」断流项 ——
 *                            换段（含首段起始）当拍置 _bSegNew，次拍 _bSegReset 为真使 IN 断流，
 *                            ET 归零后再起计，故单段超时按段独立（结构性无需外部沿清零）。
 *                         ② 斜坡双向：目标高于当前则升、低于当前则降（段间降力不越界），
 *                            三步比较全用大小判据，无浮点等值比较（R4）。
 *                         ③ 到力容差为「相对 0.5% 与绝对 0.1 kN 取大」，浮点比较一律容差式。
 *                         ④ 组态域闸：nSegCnt ∈ [1,4]（越域直接故障并钳位供下标安全）；
 *                            参与执行的段（1..nSegCnt）逐段校验速率 > 0、目标力 ≥ 0、保压 ≤ 1h；
 *                            全部 4 段做非有限拒收（未参与段不判量程域，见分工声明）。
 *                         ⑤ 无除法，故无除零；无浮点等值比较；力指令出口恒为饱和值。
 *                         ⑥ 零全局耦合（无 GVL / VAR_EXTERNAL / %I / %Q，R1 / R2）。
 * 码表     (Codes)      : 本件不占用全局数字码位（R297 零码位范式）；出口为 BOOL + ENUM，
 *                         enum E_DL_PfcPhase / E_DL_PfcCause 归属本文件（全库唯一属主，R264）。
 *                         信息级（0..9）永不置 bError；故障级（10 起）赋值处与 _bFaultLatch 三行
 *                         成对（R45），锁存回放至 bReset 沿（FB33-1）。
 * 分工声明 (Scope)      : 压机液压比例阀闭环 / 伺服压力闭环归运动控制件；模具保护与吨位监视归
 *                         FB_DL_PressTonnageGuard 类件；本件只做**多段力配方开环斜坡 + 到力判定 +
 *                         保压计时**，不做力闭环 PID，也不做安全回路（安全由 PRG_IoMapping 双切断）。
 * 归属     (Ownership)  : E_DL_PfcPhase / E_DL_PfcCause 归属本文件（全库唯一定义，R264）。
 * 红线自检 (Redline)    : R1 ✓ 零 GVL ｜ R2 ✓ 零 %I/%Q ｜ R3 ✓ 纯 IEC ｜ R4 ✓ dt 闸 + 容差比较 +
 *                         非有限双判 + 无除法 ｜ R5 ✓ 逐行同行双语注释 ｜ R6 ✓ 六态 ENUM + CASE +
 *                         ELSE ｜ R7 ✓ 全部 TON/R_TRIG 在 CASE 外 ｜ R8/R9 N/A（无 METHOD）
 *                         R10 ✓ 无构造式转换 ｜ R14 ✓ 无 PROPERTY ｜ R15 ✓ 无保留字撞名
 *                         R17 ✓ 定长 ARRAY[1..4] ｜ R18 ✓ bReset 用 R_TRIG 判 .Q ｜ R19 ✓ eFault
 *                         出口 = bReset 沿 + 撤使能 ｜ R20 ✓ 到力等待相带 tSegTimeout 超时兜底
 *                         R21 ✓ 锁存与迁相分离。
 * 修订历史 (Revision)   : 2026-11-24  v1.0.0  R79-B 首版
 * 验收向量 (Acceptance) :
 *   V1 nSegCnt=2、段1 = (50 kN, 10 kN/s, T#2S)、段2 = (80 kN, 5 kN/s, T#1S)、tSegTimeout=T#30S、
 *      fForceFb 跟随 fForceCmd：eRamp 约 5s 到 50 kN → eHold（tHoldElapsed 递增到 2s）→ 段2：
 *      约 6s 到 80 kN → eHold 1s → eRelease → eDone，bCurveDone=TRUE、nSegCompleted=2。
 *   V2 nSegCnt=0（越域）→ eState=eFault、eCause=eBadConfig、bError=TRUE、fForceCmd=0；
 *      bReset 上升沿且 bEnable=FALSE → 回 eIdle、bError=FALSE。
 *   V3 aSegRate[1]=0.0（速率非正）→ eState=eFault、eCause=eBadConfig。
 *   V4 aSegForce[1]=50.0、tSegTimeout=T#5S、fForceFb 恒为 0（力建不起来）→ 5s 后
 *      eState=eFault、eCause=eForceNotReached、bError=TRUE、fForceCmd=0（故障相全撤）。
 *   V5 fForceFb = NaN → eState=eFault、eCause=eNonFinite（非有限拒收，非量程判据）。
 *   V6 eRamp 中 bStart 落 FALSE → fForceCmd 回 0、eState=eIdle、nSegAct=0（安全降级）。
 *============================================================================*)

(*-----------------------------------------------------------------------------
 * 枚举: E_DL_PfcPhase（压机力曲线相位；eFault 为安全相，仅 bReset 沿迁出）
 *----------------------------------------------------------------------------*)
TYPE E_DL_PfcPhase :
(
    eIdle    := 0,    // 空闲：力指令 0，段号清零 / Idle: force command zero, segment cleared
    eRamp    := 10,   // 斜坡相：按段速率逼近目标力 / Ramp: approach the target at the segment rate
    eHold    := 20,   // 保压相：力保持目标值并计时 / Hold: keep the target force and time it
    eRelease := 30,   // 卸力相：力指令斜坡降到 0 / Release: ramp the force command down to zero
    eDone    := 40,   // 完成相：bCurveDone 电平为 TRUE / Done: bCurveDone held high
    eFault   := 90    // 故障安全相：锁存成因，力指令回 0 / Fault safe phase: latched cause, force command zeroed
);
END_TYPE

(*-----------------------------------------------------------------------------
 * 枚举: E_DL_PfcCause（成因码；信息级 = 0..9，故障级 = 10 起）
 *----------------------------------------------------------------------------*)
TYPE E_DL_PfcCause :
(
    eNone            := 0,   // 信息级：无事件 / Info: no event
    eSegDone         := 1,   // 信息级：一段保压完成 / Info: one segment hold completed
    eCurveDoneCode   := 2,   // 信息级：曲线保压全部完成 / Info: all segment holds completed
    eReleasing       := 3,   // 信息级：进入卸力相 / Info: entering the release phase
    eBadConfig       := 10,  // 故障级：段数 / 速率 / 目标力 / 保压 / 超时越域 / Fault: segment, rate, force, hold or timeout out of domain
    eNonFinite       := 11,  // 故障级：入参非有限 / Fault: non-finite input
    eForceNotReached := 12,  // 故障级：单段超时未到力 / Fault: force not reached within the segment timeout
    eIllegalState    := 13   // 故障级：非法状态枚举值 / Fault: illegal state enum value
);
END_TYPE

FUNCTION_BLOCK FB_DL_PressForceCurveExec
VAR_INPUT
    bEnable     : BOOL := FALSE;                        // 使能：FALSE 力指令回 0 并回 eIdle / Enable, FALSE zeroes the force and returns to idle
    bStart      : BOOL := FALSE;                        // 启动（电平）：FALSE 曲线中止，力指返回 0 / Start level, FALSE aborts and ramps the force back
    bReset      : BOOL := FALSE;                        // 复位（上升沿，需同时 bEnable=FALSE）/ Reset rising edge, requires bEnable FALSE
    aSegForce   : ARRAY[1..4] OF LREAL;                 // 各段目标力（域 ≥ 0）[kN] / Per-segment target force, domain >= 0
    aSegRate    : ARRAY[1..4] OF LREAL;                 // 各段升力速率（域 > 0）[kN/s] / Per-segment force rate, domain > 0
    aSegHold    : ARRAY[1..4] OF TIME;                  // 各段保压时长（域 0..1h）[s] / Per-segment hold time, domain 0..1h
    nSegCnt     : INT := 1;                             // 实际执行段数，有效域 1..4 [段] / Effective segment count, valid domain 1..4
    fForceFb    : LREAL := 0.0;                         // 实际力反馈（来自压力/力传感器）[kN] / Actual force feedback
    tSegTimeout : TIME := T#30S;                        // 单段到力超时，域 100ms..1h [s] / Per-segment force-reach timeout
END_VAR
VAR_OUTPUT
    fForceCmd      : LREAL := 0.0;                      // 力指令出口（斜坡饱和值）[kN] / Force command outlet, saturated ramp value
    nSegAct        : INT := 0;                          // 当前段号（1 起，0 = 未开始）[段] / Current segment number, 0 means not started
    tHoldElapsed   : TIME := T#0S;                      // 当前段保压已用时长 [s] / Elapsed hold time of the current segment
    bCurveDone     : BOOL;                              // 曲线完成（电平，保持至 bStart 落或复位）[-] / Curve done, level held until start falls
    eState         : E_DL_PfcPhase;                     // 状态出口（段尾单点映射）[-] / State outlet mapped at the tail
    eCause         : E_DL_PfcCause;                     // 成因码出口（故障期锁存回放）[-] / Cause code outlet
    bError         : BOOL;                              // 故障锁存标志 [-] / Fault latch flag
    bValid         : BOOL;                              // 曲线有效回执（斜坡/保压相且无锁存）[-] / Curve validity receipt
    nSegCompleted  : INT := 0;                          // 已完成段数 [段] / Number of completed segments
END_VAR
VAR
    _eState       : E_DL_PfcPhase := E_DL_PfcPhase.eIdle;   // 内部相位（CASE 唯一写入目标）[-] / Internal phase
    _bFaultLatch  : BOOL := FALSE;                          // 故障锁存位（仅 bReset 沿清除）[-] / Fault latch bit
    _eCauseLatch  : E_DL_PfcCause := E_DL_PfcCause.eNone;    // 锁存成因码（FB33-1 锁存回放）[-] / Latched cause code
    _eCauseTmp    : E_DL_PfcCause := E_DL_PfcCause.eNone;    // 本拍首因中间量（段 6 组态闸用）[-] / First cause of this scan
    _bCfgOk       : BOOL := TRUE;                           // 组态与入参闸通过标志 [-] / Configuration gate flag
    _bResetPulse  : BOOL := FALSE;                          // bReset 上升沿快照（R18）[-] / bReset rising-edge snapshot
    _nSegClamp    : INT := 1;                               // 段数钳位值 1..4（下标安全）[段] / Clamped segment count for safe indexing
    _bSegNew      : BOOL := FALSE;                          // 本拍进入新段标志（CASE 内置位，次拍令单段超时 ET 自清）[-] / New-segment flag set inside CASE
    _bSegReset    : BOOL := FALSE;                          // 新段标志快照（段 1 取上一拍值，供 tonSeg 的 IN 断流）[-] / New-segment snapshot latching the last-scan value
    _nIdx         : INT := 1;                               // 遍历下标（FOR 专用）[段] / Loop index for FOR statements
    _diHoldMs     : DINT := 0;                              // 保压毫秒累加（DINT 防跨型溢出）[ms] / Accumulated hold milliseconds
    _fDtSec       : LREAL := 0.0;                           // 采样步长 [s] / Sampling step in seconds
    _bDtOk        : BOOL := FALSE;                          // 步长有效性（dt > EPS）[-] / Sampling step validity
    _fStep         : LREAL := 0.0;                          // 本拍斜坡增量 [kN] / Ramp increment of this scan
    _fTol         : LREAL := 0.0;                           // 到力容差 = max(0.5%×|目标|, 0.1) [kN] / Force-reach tolerance
    _bCmdAtTarget : BOOL := FALSE;                          // 指令已饱和到目标标志 [-] / Command saturated at the target
    _bFbInTol     : BOOL := FALSE;                          // 反馈落进容差带标志 [-] / Feedback inside the tolerance band
    rtReset       : R_TRIG;                                 // bReset 边沿实例（段 4 无条件调用，R18）/ bReset edge instance called unconditionally
    tonDt         : TON;                                    // 定周期采样节拍（段 4 无条件调用）/ Fixed-period sampling tick
    tonSeg        : TON;                                    // 单段到力超时（段 4 无条件调用）/ Per-segment force-reach timeout
END_VAR
VAR CONSTANT
    DL_PFC_ZERO      : LREAL := 0.0;             // 浮点零基准 [-] / Float zero base
    DL_PFC_EPS       : LREAL := 1.0E-6;          // 浮点同值/正步长容差（力指令饱和判）[-] / Float equality and positive-step tolerance
    DL_PFC_TOL_PCT   : LREAL := 0.005;           // 到力相对容差 0.5% [-] / Relative force tolerance of 0.5 percent
    DL_PFC_TOL_ABS   : LREAL := 0.1;             // 到力绝对容差 [kN] / Absolute force tolerance
    DL_PFC_SEG_MAX   : INT := 4;                 // 段数上限（数组定长）[段] / Upper bound of segments, fixed array size
    DL_PFC_ONE       : INT := 1;                 // 段号起始值 [段] / Segment numbering start
    DL_PFC_DT        : TIME := T#100MS;          // 采样节拍（斜坡步长来源）[s] / Sampling tick, the ramp step source
    DL_PFC_DT_MS     : DINT := 100;              // 采样节拍毫秒数（保压累加步长）[ms] / Sampling tick in milliseconds
    DL_PFC_T_MIN     : TIME := T#100MS;          // 超时参数下限 [s] / Lower bound of the timeout parameter
    DL_PFC_T_MAX     : TIME := T#1H;             // 超时与保压参数上限 [s] / Upper bound of timeout and hold time
    DL_PFC_MS_ZERO   : DINT := 0;                // 毫秒零基准 [-] / Millisecond zero base
END_VAR

(* —— 段 1：单拍与电平出口预置（不清锁存 / 力指令 / 段号状态，FB32-1） —— *)
bCurveDone := FALSE;                                   // 曲线完成电平每拍预清（仅 eDone 相重新置位）/ Curve-done level preset, re-armed only in eDone
_bCfgOk    := TRUE;                                    // 组态闸标志复位 / Configuration flag reset
_eCauseTmp := E_DL_PfcCause.eNone;                      // 当拍首因复位 / Scan cause reset
_bSegReset := _bSegNew;                                // 取上一拍的新段标志（本拍令 tonSeg 的 IN 断流，R188）/ Take the last-scan new-segment flag
_bSegNew   := FALSE;                                   // 新段标志每拍预清（仅换段相内置位）/ Preset the new-segment flag, set only on a segment change

(* —— 段 2：段数钳位与采样步长（标准转换，R10） —— *)
_nSegClamp := LIMIT(DL_PFC_ONE, nSegCnt, DL_PFC_SEG_MAX);            // 段数钳位 1..4 / Clamp the segment count
_fDtSec    := TIME_TO_LREAL(DL_PFC_DT);                              // 节拍换算为秒 / Sampling tick to seconds
IF _fDtSec > DL_PFC_EPS THEN
    _bDtOk := TRUE;                                                  // 步长为正：允许斜坡积分 / Positive step: ramp integration allowed
ELSE
    _bDtOk := FALSE;                                                 // 步长非正：拒绝积分（R4）/ Non-positive step: integration refused
END_IF

(* —— 段 3：全部 4 段非有限拒收（未参与段也拒 NaN / Inf，避免污染后续组态）/ —— *)
FOR _nIdx := 1 TO DL_PFC_SEG_MAX DO
    IF (aSegForce[_nIdx] <> aSegForce[_nIdx]) OR ((aSegForce[_nIdx] - aSegForce[_nIdx]) <> DL_PFC_ZERO) THEN
        _bCfgOk    := FALSE;                            // 目标力非有限 / Target force is not finite
        _eCauseTmp := E_DL_PfcCause.eNonFinite;         // 故障级：非有限入参 / Fault: non-finite input
    END_IF
    IF (aSegRate[_nIdx] <> aSegRate[_nIdx]) OR ((aSegRate[_nIdx] - aSegRate[_nIdx]) <> DL_PFC_ZERO) THEN
        _bCfgOk    := FALSE;                            // 速率非有限 / Rate is not finite
        _eCauseTmp := E_DL_PfcCause.eNonFinite;         // 故障级：非有限入参 / Fault: non-finite input
    END_IF
END_FOR
IF (fForceFb <> fForceFb) OR ((fForceFb - fForceFb) <> DL_PFC_ZERO) THEN
    _bCfgOk    := FALSE;                                // 力反馈非有限 / Force feedback is not finite
    _eCauseTmp := E_DL_PfcCause.eNonFinite;             // 故障级：非有限入参 / Fault: non-finite input
END_IF

(* —— 段 4：组态量程域闸（仅参与执行的 1..nSegCnt 段，逐段校验） —— *)
IF _bCfgOk THEN
    IF (nSegCnt < DL_PFC_ONE) OR (nSegCnt > DL_PFC_SEG_MAX) THEN
        _bCfgOk    := FALSE;                            // 段数越域 / Segment count out of domain
        _eCauseTmp := E_DL_PfcCause.eBadConfig;         // 故障级：组态非法 / Fault: bad configuration
    ELSIF (tSegTimeout < DL_PFC_T_MIN) OR (tSegTimeout > DL_PFC_T_MAX) THEN
        _bCfgOk    := FALSE;                            // 单段超时越域 / Segment timeout out of domain
        _eCauseTmp := E_DL_PfcCause.eBadConfig;         // 故障级：组态非法 / Fault: bad configuration
    ELSE
        FOR _nIdx := 1 TO _nSegClamp DO
            IF aSegRate[_nIdx] <= DL_PFC_ZERO THEN
                _bCfgOk    := FALSE;                    // 速率非正，无法斜坡 / Non-positive rate, ramp impossible
                _eCauseTmp := E_DL_PfcCause.eBadConfig; // 故障级：组态非法 / Fault: bad configuration
            END_IF
            IF aSegForce[_nIdx] < DL_PFC_ZERO THEN
                _bCfgOk    := FALSE;                    // 目标力为负 / Negative target force
                _eCauseTmp := E_DL_PfcCause.eBadConfig; // 故障级：组态非法 / Fault: bad configuration
            END_IF
            IF aSegHold[_nIdx] > DL_PFC_T_MAX THEN
                _bCfgOk    := FALSE;                    // 保压时长越上限 / Hold time above the upper bound
                _eCauseTmp := E_DL_PfcCause.eBadConfig; // 故障级：组态非法 / Fault: bad configuration
            END_IF
        END_FOR
    END_IF
END_IF

(* —— 段 5：边沿与定时器（CASE 外无条件调用，R7；IN 均含 NOT .Q 自复位，R188） —— *)
rtReset(CLK := bReset);                                // bReset 边沿无条件刷新（R18）/ bReset edge refreshed unconditionally
_bResetPulse := rtReset.Q;                             // 边沿快照 / Edge snapshot
tonDt(IN := ((_eState = E_DL_PfcPhase.eRamp) OR (_eState = E_DL_PfcPhase.eHold)
             OR (_eState = E_DL_PfcPhase.eRelease))
            AND (NOT tonDt.Q) AND (NOT _bFaultLatch),
      PT := DL_PFC_DT);                                // 执行相定周期采样节拍 / Fixed-period tick in the execution phases
tonSeg(IN := (_eState = E_DL_PfcPhase.eRamp) AND (NOT _bSegReset)
              AND (NOT tonSeg.Q) AND (NOT _bFaultLatch),
        PT := tSegTimeout);                            // 单段超时：换段次拍 IN 断流使 ET 自清（R188）

(* —— 段 6：状态机主体（唯一相位写入点；故障只置锁存，迁相由段 8 统一执行） —— *)
CASE _eState OF
    E_DL_PfcPhase.eIdle :
        fForceCmd     := DL_PFC_ZERO;                  // 空闲：力指令归零 / Idle: force command zeroed
        nSegAct       := 0;                            // 空闲：段号清零 / Idle: segment cleared
        nSegCompleted := 0;                            // 空闲：完成段数清零 / Idle: completed segments cleared
        _diHoldMs     := DL_PFC_MS_ZERO;               // 空闲：保压累计清零 / Idle: hold accumulator cleared
        IF bEnable AND bStart AND _bCfgOk AND (NOT _bFaultLatch) THEN
            fForceCmd  := DL_PFC_ZERO;                 // 迁移①：起点力为零 / Start from zero force
            nSegAct    := DL_PFC_ONE;                  // 从第 1 段开始 / Begin at segment one
            _diHoldMs  := DL_PFC_MS_ZERO;              // 保压累计清零 / Hold accumulator cleared
            _bSegNew   := TRUE;                        // 首段起始：次拍令单段超时 ET 自清 / First segment: reset the timeout on the next scan
            eCause     := E_DL_PfcCause.eNone;         // 信息级：无事件 / Info: no event
            _eState    := E_DL_PfcPhase.eRamp;         // 进入斜坡相 / Move to ramp
        END_IF

    E_DL_PfcPhase.eRamp :
        IF (NOT bEnable) OR (NOT bStart) THEN
            fForceCmd := DL_PFC_ZERO;                  // 失能：力指令回 0（安全降级）/ Disabled: force zeroed for safety
            nSegAct   := 0;                            // 段号清零 / Segment cleared
            eCause    := E_DL_PfcCause.eNone;          // 信息级：无事件 / Info: no event
            _eState   := E_DL_PfcPhase.eIdle;          // 回空闲相 / Back to idle
        ELSE
            (* 斜坡：按段速率把力指令推向目标（双向） *)
            IF tonDt.Q AND _bDtOk THEN
                _fStep := aSegRate[nSegAct] * _fDtSec; // 本拍增量 = 速率 × dt [kN]
                IF fForceCmd < aSegForce[nSegAct] THEN
                    fForceCmd := MIN(fForceCmd + _fStep, aSegForce[nSegAct]);   // 升力且不越过目标 / Ramp up without overshoot
                ELSIF fForceCmd > aSegForce[nSegAct] THEN
                    fForceCmd := MAX(fForceCmd - _fStep, aSegForce[nSegAct]);   // 降力且不越过目标 / Ramp down without overshoot
                END_IF
            END_IF
            (* 到力判据：容差 = max(0.5%×|目标|, 0.1 kN)，浮点比较一律容差式（R4） *)
            _fTol := MAX(ABS(aSegForce[nSegAct]) * DL_PFC_TOL_PCT, DL_PFC_TOL_ABS);
            _bCmdAtTarget := ABS(fForceCmd - aSegForce[nSegAct]) <= DL_PFC_EPS;   // 指令已饱和到目标
            _bFbInTol     := ABS(fForceFb - aSegForce[nSegAct]) <= _fTol;         // 反馈落进容差带
            IF _bCmdAtTarget AND _bFbInTol THEN
                fForceCmd := aSegForce[nSegAct];       // 迁移②：到力，指令精确取目标 / Reached: command set exactly
                _diHoldMs := DL_PFC_MS_ZERO;           // 保压累计清零 / Hold accumulator cleared
                eCause    := E_DL_PfcCause.eNone;      // 信息级：无事件 / Info: no event
                _eState   := E_DL_PfcPhase.eHold;      // 进入保压相 / Move to hold
            ELSIF tonSeg.Q THEN
                IF NOT _bFaultLatch THEN
                    _eCauseLatch := E_DL_PfcCause.eForceNotReached;   // 故障级：单段超时未到力 / Fault: force not reached
                    _bFaultLatch := TRUE;                             // 置故障锁存（迁相由段 8，R21）/ Latch the fault
                END_IF
            END_IF
        END_IF

    E_DL_PfcPhase.eHold :
        IF (NOT bEnable) OR (NOT bStart) THEN
            fForceCmd := DL_PFC_ZERO;                  // 失能：力指令回 0 / Disabled: force zeroed
            nSegAct   := 0;                            // 段号清零 / Segment cleared
            eCause    := E_DL_PfcCause.eNone;          // 信息级：无事件 / Info: no event
            _eState   := E_DL_PfcPhase.eIdle;          // 回空闲相 / Back to idle
        ELSE
            fForceCmd := aSegForce[nSegAct];           // 保压相：力指令锁定目标值 / Hold: command locked to the target
            IF tonDt.Q AND _bDtOk THEN
                _diHoldMs := _diHoldMs + DL_PFC_DT_MS; // 保压毫秒累加 / Accumulate hold milliseconds
            END_IF
            IF _diHoldMs >= TIME_TO_DINT(aSegHold[nSegAct]) THEN
                nSegCompleted := nSegCompleted + DL_PFC_ONE;   // 本段完成计数 / Count the completed segment
                _diHoldMs     := DL_PFC_MS_ZERO;               // 保压累计清零 / Hold accumulator cleared
                IF nSegAct >= _nSegClamp THEN
                    eCause  := E_DL_PfcCause.eCurveDoneCode;    // 迁移④：末段完成 / Info: last segment done
                    _eState := E_DL_PfcPhase.eRelease;          // 进入卸力相 / Move to release
                ELSE
                    nSegAct := nSegAct + DL_PFC_ONE;            // 迁移③：进入下一段 / Next segment
                    _bSegNew := TRUE;                           // 换段：次拍令单段超时 ET 自清 / Segment change: reset the timeout next scan
                    eCause  := E_DL_PfcCause.eSegDone;          // 信息级：一段完成 / Info: one segment done
                    _eState := E_DL_PfcPhase.eRamp;             // 回斜坡相 / Back to ramp
                END_IF
            END_IF
        END_IF

    E_DL_PfcPhase.eRelease :
        IF (NOT bEnable) OR (NOT bStart) THEN
            fForceCmd := DL_PFC_ZERO;                  // 失能：力指令直接归零 / Disabled: force zeroed immediately
            nSegAct   := 0;                            // 段号清零 / Segment cleared
            eCause    := E_DL_PfcCause.eNone;          // 信息级：无事件 / Info: no event
            _eState   := E_DL_PfcPhase.eIdle;          // 回空闲相 / Back to idle
        ELSE
            eCause := E_DL_PfcCause.eReleasing;        // 信息级：卸力中 / Info: releasing
            IF tonDt.Q AND _bDtOk THEN
                _fStep := aSegRate[_nSegClamp] * _fDtSec;                  // 卸力速率取末段速率 / Release rate from the last segment
                fForceCmd := fForceCmd - _fStep;                           // 力指令斜坡下降 / Ramp the command down
                IF fForceCmd < DL_PFC_ZERO THEN
                    fForceCmd := DL_PFC_ZERO;                              // 下限饱和，防负力指令 / Clamp at zero, no negative command
                END_IF
            END_IF
            IF ABS(fForceCmd) <= DL_PFC_EPS THEN
                fForceCmd := DL_PFC_ZERO;              // 迁移⑤：已退到 0，精确归零 / Fully released: exact zero
                eCause    := E_DL_PfcCause.eCurveDoneCode;   // 信息级：曲线完成 / Info: curve completed
                _eState   := E_DL_PfcPhase.eDone;      // 进入完成相 / Move to done
            END_IF
        END_IF

    E_DL_PfcPhase.eDone :
        fForceCmd  := DL_PFC_ZERO;                     // 完成相：力指令保持 0 / Done: force stays zero
        bCurveDone := TRUE;                            // 曲线完成电平 / Curve-done level high
        IF (NOT bStart) OR _bResetPulse THEN
            bCurveDone    := FALSE;                    // 迁移⑥：撤完成电平 / Withdraw the done level
            nSegAct       := 0;                        // 段号清零 / Segment cleared
            nSegCompleted := 0;                        // 完成段数清零 / Completed segments cleared
            eCause        := E_DL_PfcCause.eNone;      // 信息级：无事件 / Info: no event
            _eState       := E_DL_PfcPhase.eIdle;      // 回空闲相 / Back to idle
        END_IF

    E_DL_PfcPhase.eFault :
        fForceCmd := DL_PFC_ZERO;                      // 故障相：力指令回 0（安全侧）/ Fault phase: force zeroed
        IF _bResetPulse AND (NOT bEnable) THEN
            _bFaultLatch  := FALSE;                    // 迁移⑨：清故障锁存 / Clear the fault latch
            _eCauseLatch  := E_DL_PfcCause.eNone;      // 清锁存成因 / Clear the latched cause
            eCause        := E_DL_PfcCause.eNone;      // 出口同步归零 / Outlet follows
            nSegAct       := 0;                        // 段号清零 / Segment cleared
            nSegCompleted := 0;                        // 完成段数清零 / Completed segments cleared
            _diHoldMs     := DL_PFC_MS_ZERO;           // 保压累计清零 / Hold accumulator cleared
            _eState       := E_DL_PfcPhase.eIdle;      // 回空闲相 / Back to idle
        END_IF

ELSE
    (* 迁移⑩：非法枚举兜底（R6） *)
    IF NOT _bFaultLatch THEN
        _eCauseLatch := E_DL_PfcCause.eIllegalState;   // 故障级：非法状态 / Fault: illegal state
        _bFaultLatch := TRUE;                          // 置故障锁存 / Latch the fault
    END_IF
END_CASE

(* —— 段 7：组态闸失败处理（锁存与迁相分离，R21） —— *)
IF (NOT _bCfgOk) AND (NOT _bFaultLatch) THEN
    _eCauseLatch := _eCauseTmp;                        // 锁存首因（组态闸）/ Latch the configuration cause
    _bFaultLatch := TRUE;                              // 置故障锁存 / Latch the fault
END_IF

(* —— 段 8：段尾故障迁移闸 + 故障相动作全撤（FB50-1④） —— *)
IF _bFaultLatch AND (_eState <> E_DL_PfcPhase.eFault) THEN
    _eState := E_DL_PfcPhase.eFault;                   // 锁存即迁相 / Latch forces the fault phase
END_IF
IF _eState = E_DL_PfcPhase.eFault THEN
    fForceCmd  := DL_PFC_ZERO;                         // 故障相力指令全撤（含同拍迁入）/ Force withdrawn in fault
    bCurveDone := FALSE;                               // 故障相撤完成电平 / Done level withdrawn in fault
END_IF

(* —— 段 9：统一出口（状态映射 + 保压时长换算 + 锁存回放） —— *)
eState       := _eState;                               // 相位映射 / Phase mapping
tHoldElapsed := DINT_TO_TIME(_diHoldMs);               // 保压毫秒 → TIME（标准转换）/ Hold milliseconds to TIME
bError       := _bFaultLatch;                          // 故障标志取锁存位 / Fault flag from the latch
IF _bFaultLatch THEN
    eCause := _eCauseLatch;                            // 故障期回放锁存码（FB33-1）/ Replay the latched code
END_IF
bValid := ((_eState = E_DL_PfcPhase.eRamp) OR (_eState = E_DL_PfcPhase.eHold)
           OR (_eState = E_DL_PfcPhase.eRelease)) AND (NOT _bFaultLatch);   // 执行相且无锁存时有效
END_FUNCTION_BLOCK

(* ---- FB_DL_ReactorJacketDeltaT.st ---- *)
(*==============================================================================
 * 组件名称 (Component)  : FB_DL_ReactorJacketDeltaT
 * 所属子库 (Sublibrary) : DL_Process
 * 当前版本 (Version)    : 1.0.0
 * 组件分类 (Category)   : 功能块（FUNCTION_BLOCK）· 釜温-夹套温差约束与冷热分程
 * 兼容性   (Platform)   : CODESYS 3.5 / TwinCAT 3 / 汇川 InoProShop / Schneider Machine Expert
 *                         仅依赖 Standard.library（R_TRIG / TON / ABS / MIN / MAX / LIMIT）
 *                         与库内低层件 FB_DL_RateLimiter（DL_Algo），零厂商方言
 * 接口依赖 (Depends)    : E_DL_Ne107Status（属主 A1）、FB_DL_RateLimiter（DL_Algo 既有件）。
 *                         温度闭环由 FB_DL_CascadePid 承担，本件只做「约束层 + 分程层」。
 * 功能描述 (Function)   : 放热反应的釜温-夹套温差抑制。以 ΔT = 釜温 − 夹套温 为约束量，
 *                         对升温侧做**温差上限约束**与**温差变化率约束**，并把上层 PID 输出
 *                         分程为冷/热两路阀位给定；超温时强制冷却；分程带死区防冷热同开。
 * 边界与纪律 (Boundary) : ① **不内联 PID** —— 温度闭环由 FB_DL_CascadePid 承担，PID 输出以
 *                         fPidOut 引脚注入，本件绝不实现比例/积分/微分；② **不新增轴/相状态
 *                         枚举** —— 工艺相状态归 FB_DL_BatchPhaseBase，本件的 E_DL_JacketState
 *                         只描述「冷热分程的当前执行方向」，不是批次相状态（R31 家族纪律）；
 *                         ③ 两路输出**互斥**（由状态机与目标量赋值保证），并带 fDeadband 死区，
 *                         禁止「冷热同开」；④ 不做阀位反馈校验（归阀门件）。
 * 分层声明 (Layer)      : 工艺层（DL_Process）。限速能力**组合调用** FB_DL_RateLimiter，
 *                         绝不内联限速算法（依赖方向纪律）。零全局变量表引用、零外部变量声明、
 *                         零物理 IO 地址。
 * 段序     (Segments)   : 段1 实例无条件刷新（含两个限速器实例）→ 段2 复位通道（CASE 前，R39）→
 *                         段3 输入防御与参数钳位 → 段4 温差与变化率测量（TON 统计窗，R40）→
 *                         段5 状态机（约束层 + 分程层）→ 段6 分程限速（组合低层件）→
 *                         段7 码位单一优先级链 → 段8 出口钳位与互斥仲裁。
 * 枚举映射表 (R31)      : eIdle(0)→标签 0｜eHeat(10)→标签 10｜eCool(20)→标签 20｜eHold(30)→标签 30｜
 *                         eFault(99)→标签 99。每个成员有且仅有一个显式标签，ELSE 只接脏值（02FE）。
 * 单拍标志清单 (R25)    : 本件唯一的沿输入是 bReset：预清零点段1 每拍覆盖 _bResetEdge；置位点
 *                         段1 的 _fbTrigReset 实例调用；自清点紧随实例调用的赋值行。
 * 保持位清单 (R27)      : bDeltaTLimited / bOverTemp / fHeatOut / fCoolOut —— 逐拍由
 *                         _bLimitLatched / _bOverTempLatched / 限速器输出重写，绝不靠进入那拍。
 * 定时器清单 (R40)      : _fbTonRate｜IN = NOT _bRateBreak（变化率统计窗，PT = tRateWindow）｜
 *                         断输入标志 _bRateBreak（每次窗口结算置一拍，ET 归零后重开新窗）｜
 *                         自清点：段2 无条件 `IF _bRateBreak THEN _bRateBreak := FALSE; END_IF`。
 *                         另有两个 FB_DL_RateLimiter 实例在段6 无条件周期调用（R7：位于主体顶层，
 *                         不在任何 IF/CASE 之内；必须在状态机算出目标量之后，否则目标滞后一拍）。
 * 三元一致表 (R35)      : 温差上限守卫 5~150 K / 封顶 150 / 判据 `>=`（达上限即冻结）｜
 *                         变化率守卫 0.1~50 K/min / 封顶 50 / 判据 `>`（超阈只报警不拦截）｜
 *                         死区守卫 0~10 % / 封顶 10 / 判据 `<=`（判据 `<=` 与封顶同向）。
 * 镜像量清单 (R38)      : fReactorTemp / fJacketTemp / fPidOut 的唯一消费点是段3 的三个快照
 *                         （_fReactorNow / _fJacketNow / _fPidNow），全件不二次读取实时入参。
 * R36 关联（必须手算，写给调用方）: 本件消费上层 PID 输出 fPidOut。**调用方须保证 fPidOut 已过
 *                         「跟踪结束首拍」处理**：若上层 PID 处于跟踪态（手动/暂停）时输出为
 *                         fTrack，切自动首拍 fPidOut = fP + fI + fD 可能相对 fTrack 跳变
 *                         Δ = fPidOut − fTrack。手算示例：fTrack = 0 %、fP = 24 %、fI = 18 %、
 *                         fD = 0 %（微分先行且无扰动）→ 首拍 fPidOut = 42 %，跳变 42 %；若上层
 *                         PID 已按无扰切换（fI := fOut − fP − fD 反算残量）则 fI 已被重算为
 *                         −24 %，首拍 fPidOut 仍为 0 %，不会出现阶跃。本件对该阶跃**不做补偿**
 *                         （补偿属 PID 的无扰切换职责），只保证：首拍大跳不会触发 16#0005_01CF
 *                         （01CF 的判据是实测温差达上限，不是指令跳变）。V4 向量复现该场景。
 * 开源溯源 (Origin)     : 原创实现（参考 Siemens LBP 的「给定 → 限幅 → 闭环 → 执行机构限幅」
 *                         设定值分层组织结构，T2-2 主源；以及 ISA-88 公开的相语义与状态迁移
 *                         惯例，T2-8 次源）。仅借分层骨架与参数域划分，LBP 块名、参数名、UDT
 *                         布局、门限值一律未沿用；温差约束、分程死区、反装判据为本库自有。
 *                         许可证说明：LBP 与 ISA-88 均为文档/公开规范（非代码），只借组织
 *                         结构，clean-room 编写；本文件为本库原创，随本库许可证发布。
 * 验收向量 (Acceptance) :
 *   V1 釜 80 ℃、夹套 60 ℃、fPidOut = +40 %、fDeltaTMax = 30 → eHeat、fHeatOut = 40.0、
 *      fCoolOut = 0.0（未受限时不限速，直接跟随）。
 *   V2（约束层）釜温继续升、ΔT = 31 K → bDeltaTLimited = TRUE、fHeatOut 按 fDeltaTRate
 *      折算的速率斜坡回 0、16#0005_01CF。
 *   V3（V-C 死区分程）fPidOut = +1.0 %（< 死区 2.0）→ 两路均 0（eHold），**不得**冷热同开；
 *      离开死区时置 16#0005_01D1。
 *   V4（V-D R36 跟踪首拍）上层 PID 从手动跟踪切自动，首拍 fPidOut 由 0 跳到 +60 % → 本件
 *      未受限时直通（周期内不产生 ΔT 变化），**不得**因此误报 01CF；一旦因温差触限，输出按
 *      fDeltaTRate 限速回落（限速路径由 FB_DL_RateLimiter 承担，非限幅）。
 *   V5（V-A 反装）釜 80、夹套 95、fPidOut = +50 % → ΔT = −15 且要求升温 → 16#0005_02FD 锁存
 *      （这是本件最有价值的一条：反装传感器会被这条抓住）。
 * 偏离留档 (Deviation)  :
 *   ① 增补 tCycle 引脚（任务扫描周期）：FB_DL_RateLimiter 的限速步长必须用真实周期折算，
 *      规格未给该引脚。理由：公共约定（时间换算基准由引脚给）与泳道内 FB_DL_LeakTestStation
 *      先例一致，属公共约定强制项，非语义偏离。
 *   ② 常态是否限速的裁定：V1 要求「fPidOut = +40 % → fHeatOut = 40.0」，V4 要求「阶跃时限速」。
 *      两者只在「未受限」与「已受限」两种工况下并存，故本件把限速施加于**约束路径**
 *      （温差触限、超温强制冷却、以及从约束态恢复的整个过程），未受限时按 V1 直通。
 *      实现上用 FB_DL_RateLimiter 的 bTrack 引脚完成无扰切换：跟踪时输出等于输入，退出跟踪
 *      那一拍从当前值开始限速，不存在回跳。
 *   ③ 温差→阀位速率折算：以常量 DL_JKT_K_PER_PCT（默认 0.5 K/%）把 fDeltaTRate [K/min]
 *      折算为 [%/s]，即 (fDeltaTRate / 60) / DL_JKT_K_PER_PCT。该常量是夹套传热增益的
 *      工艺整定值，由调用方按装置实测整定；折算关系在头注释显式披露，不做隐藏假设。
 *   ④ 控制码 01CE 的修正：规格 V2 正文写作 01CE，但码位表把「温差达上限冻结」定为
 *      16#0005_01CF，且 01CE 已被 C5 占用（配方名截断）。本件按**码位表**执行（01CF），
 *      避免跨件撞号，此处留档。
 * 修订历史 (Revision)   :
 *   2026-11-15  v1.0.0  首版入库（Round 13 · 泳道 C · DL_Process 第 26 件）
 *============================================================================*)

(*-----------------------------------------------------------------------------
 * 枚举: E_DL_JacketState（归属 FB_DL_ReactorJacketDeltaT，同文件发布）
 * 说明: 只表达「冷热分程的当前执行方向」，**不是**批次相状态（相状态归 FB_DL_BatchPhaseBase）。
 *----------------------------------------------------------------------------*)
TYPE E_DL_JacketState :
(
    eIdle  := 0,    // 空闲：未使能或参数未就绪 / Idle, disabled or parameters not ready
    eHeat  := 10,   // 升温：热路给给定，冷路 0 / Heating, heat path commanded, cool path zero
    eCool  := 20,   // 冷却：冷路给给定，热路 0 / Cooling, cool path commanded, heat path zero
    eHold  := 30,   // 保持：两路均 0（死区内或温差触限冻结）/ Hold, both paths zero
    eFault := 99    // 故障：非有限、反装或非法状态 / Fault, non-finite, reversed sensor or illegal state
) UINT;
END_TYPE

FUNCTION_BLOCK FB_DL_ReactorJacketDeltaT
VAR_INPUT
    bEnable        : BOOL;                  // 使能（Enable），FALSE = 两路归零并回空闲；复位通道不受其屏蔽 / Enable, FALSE zeroes both paths
    bReset         : BOOL;                  // 复位（Reset），上升沿清故障与保持位 / Rising edge clears the fault and the held flags
    fReactorTemp   : REAL;                  // 釜温（Reactor temperature）[℃]，域 −50~400 / Reactor temperature [degC]
    fJacketTemp    : REAL;                  // 夹套温度（Jacket temperature）[℃]，域 −50~400 / Jacket temperature [degC]
    fPidOut        : REAL;                  // 上层 PID 输出（PID output）[%]，域 −100~100，**须已过跟踪首拍**（R36）/ PID output [%], must have passed its tracking-exit scan
    fDeltaTMax     : REAL := 30.0;          // 允许最大温差（Max allowed delta-T）[K]，域 5~150，默认 30.0 / Max allowed delta-T [K]
    fDeltaTRate    : REAL := 5.0;           // 温差变化率上限（Delta-T rate limit）[K/min]，域 0.1~50，默认 5.0 / Delta-T rate limit [K/min]
    fOverTempMargin : REAL := 5.0;          // 超温强制冷却裕量（Over-temperature margin）[K]，域 0.5~50，默认 5.0 / Over-temperature margin [K]
    fTempSetpoint  : REAL;                  // 釜温设定（Reactor setpoint）[℃]，域 −50~400，超温判据用 / Reactor setpoint [degC]
    tRateWindow    : TIME := T#1M;          // 变化率统计窗（Rate window），域 5 s~10 min，默认 1 min / Rate window
    fDeadband      : REAL := 2.0;           // 冷热分程死区（Split-range deadband）[%]，域 0~10，默认 2.0 / Split-range deadband [%]
    fOutMin        : REAL := 0.0;           // 输出下限（Output lower limit）[%]，默认 0.0 / Output lower limit [%]
    fOutMax        : REAL := 100.0;         // 输出上限（Output upper limit）[%]，默认 100.0 / Output upper limit [%]
    tCycle         : TIME := T#10MS;        // 任务扫描周期（Task cycle time）[ms]，限速步长折算基准（偏离留档①）/ Task cycle time [ms]
END_VAR

VAR_OUTPUT
    fHeatOut       : REAL;                  // 热路阀位给定（Heat output）[%]，0~100，保持语义 / Heat valve command [%], held
    fCoolOut       : REAL;                  // 冷路阀位给定（Cool output）[%]，0~100，保持语义 / Cool valve command [%], held
    fDeltaT        : REAL;                  // 实测温差（Measured delta-T）[K]，有符号 = 釜温 − 夹套温 / Measured delta-T [K], signed
    fDeltaTRateMeas : REAL;                 // 实测温差变化率（Measured delta-T rate）[K/min]，窗内斜率 / Measured delta-T rate [K/min]
    bDeltaTLimited : BOOL;                  // 温差达上限、升温侧被限（Delta-T limiting active），保持语义 / TRUE while the delta-T limit is active
    bOverTemp      : BOOL;                  // 釜温超设定加裕量（Over temperature），保持语义 / TRUE while over temperature
    eVerdict       : E_DL_JacketState;      // 当前执行方向（Verdict state），逐拍重写 / Current actuation direction, rewritten every scan
    eHealth        : E_DL_Ne107Status;      // 健康态（NE107 health），引用属主 A1 的枚举 / NE107 health, owned by A1
    uDiagCode      : UDINT;                 // 诊断码（Diagnostic code），本拍单一优先级链输出 / Diagnostic code, single priority chain
    uErrorId       : UDINT;                 // 故障码（Error code），仅故障级码，0 = 无故障 / Fault-level code, 0 = no fault
    bError         : BOOL;                  // 故障标志（Error），仅故障级码置位 / TRUE only for fault-level codes
END_VAR

VAR
    _eState        : E_DL_JacketState := E_DL_JacketState.eIdle;    // 内部状态（Internal state）/ Internal state value
    _bResetEdge    : BOOL;                  // 复位沿单拍标志（Reset one-shot flag）/ Reset one-shot flag
    _bRateBreak    : BOOL;                  // 统计窗断输入拍（Rate window break）/ Rate window break
    _uFaultCode    : UDINT;                 // 本拍故障级码（Fault-level code this scan）/ Fault-level code of this scan
    _uFaultLatched : UDINT;                 // 故障码锁存（Latched fault code），仅复位清除 / Latched fault code, reset only
    _uInfoCode     : UDINT;                 // 本拍信息级码（Info-level code this scan）/ Info-level code of this scan
    _bFaultCond    : BOOL;                  // 故障条件（Fault condition）/ Fault condition flag
    _fReactorNow   : REAL;                  // 釜温快照（Reactor temperature snapshot）[℃]，单次锁存（R38）/ Reactor snapshot [degC]
    _fJacketNow    : REAL;                  // 夹套温快照（Jacket temperature snapshot）[℃]，单次锁存（R38）/ Jacket snapshot [degC]
    _fPidNow       : REAL;                  // PID 输出快照（PID output snapshot）[%]，单次锁存（R38）/ PID snapshot [%]
    _fDeltaTMaxEff : REAL;                  // 生效温差上限（Effective delta-T limit）[K] / Effective delta-T limit [K]
    _fRateLimEff   : REAL;                  // 生效变化率上限（Effective rate limit）[K/min] / Effective rate limit [K/min]
    _fOtMarginEff  : REAL;                  // 生效超温裕量（Effective over-temp margin）[K] / Effective over-temp margin [K]
    _fDeadbandEff  : REAL;                  // 生效死区（Effective deadband）[%] / Effective deadband [%]
    _fOutLowEff    : REAL;                  // 生效输出下限（Effective output low）[%] / Effective output low [%]
    _fOutHighEff   : REAL;                  // 生效输出上限（Effective output high）[%] / Effective output high [%]
    _fRatePctS     : REAL;                  // 折算后的阀位速率（Output rate）[%/s]，偏离留档③ / Output rate [%/s]
    _fSwapTmp      : REAL;                  // 交换临时量（Swap scratch）[EU] / Swap scratch [EU]
    _fRateMin      : REAL;                  // 统计窗分钟值（Window minutes）[min] / Rate window in minutes [min]
    _fDtWinStart   : REAL;                  // 窗起点温差（Delta-T at the window start）[K] / Delta-T at the window start [K]
    _bRateInit     : BOOL;                  // 变化率窗首扫标志（Rate window first-scan flag），初值 FALSE（R19）/ Rate window init flag
    _fRateMeasInt  : REAL;                  // 内部变化率（Internal rate）[K/min] / Internal rate [K/min]
    _fHeatTgt      : REAL;                  // 热路目标（Heat target）[%]，送限速器 / Heat target [%] fed to the limiter
    _fCoolTgt      : REAL;                  // 冷路目标（Cool target）[%]，送限速器 / Cool target [%] fed to the limiter
    _bLimitActive  : BOOL;                  // 本拍处于约束路径（Limiting path active this scan）/ Limiting path active
    _bLimitLatched : BOOL;                  // 温差触限锁存（Delta-T limit latch）/ Delta-T limit latch
    _bOverTempLatched : BOOL;               // 超温锁存（Over-temperature latch）/ Over-temperature latch
    _fHeatPrev     : REAL;                  // 上一拍热路输出（Previous heat output）[%] / Previous heat output [%]
    _fCoolPrev     : REAL;                  // 上一拍冷路输出（Previous cool output）[%] / Previous cool output [%]
    _fbTrigReset   : R_TRIG;                // 复位上升沿（Reset rising edge）/ Reset rising edge
    _fbTonRate     : TON;                   // 变化率统计窗（Rate window timer）/ Rate window timer
    _fbRlHeat      : FB_DL_RateLimiter;     // 热路限速器（Heat rate limiter，组合调用低层件）/ Heat rate limiter, composed from DL_Algo
    _fbRlCool      : FB_DL_RateLimiter;     // 冷路限速器（Cool rate limiter，组合调用低层件）/ Cool rate limiter, composed from DL_Algo
END_VAR

VAR CONSTANT
    DL_JKT_REAL_MAX : REAL := 3.4E38;       // 单精度有限值判据幅值（Finite magnitude bound）/ Finite bound for REAL inputs
    DL_JKT_EPS      : REAL := 1.0E-6;       // 浮点防零容差（Divide-guard epsilon）/ Float divide-guard epsilon
    DL_JKT_TEMP_MIN : REAL := -50.0;        // 温度域下限（Temperature lower domain）[℃] / Temperature lower domain [degC]
    DL_JKT_TEMP_MAX : REAL := 400.0;        // 温度域上限（Temperature upper domain）[℃] / Temperature upper domain [degC]
    DL_JKT_PID_MAX  : REAL := 100.0;        // PID 输出域（PID output domain）[%] / PID output domain [%]
    DL_JKT_DT_LO    : REAL := 5.0;          // 温差上限域下限（Delta-T upper clamp low）[K] / Delta-T upper clamp low [K]
    DL_JKT_DT_HI    : REAL := 150.0;        // 温差上限域上限（Delta-T upper clamp high）[K] / Delta-T upper clamp high [K]
    DL_JKT_RATE_LO  : REAL := 0.1;          // 变化率域下限（Rate lower clamp）[K/min] / Rate lower clamp [K/min]
    DL_JKT_RATE_HI  : REAL := 50.0;                // 变化率域上限（Rate upper clamp）[K/min] / Rate upper clamp [K/min]
    DL_JKT_OT_LO    : REAL := 0.5;          // 超温裕量域下限（Margin lower clamp）[K] / Margin lower clamp [K]
    DL_JKT_OT_HI    : REAL := 50.0;                // 超温裕量域上限（Margin upper clamp）[K] / Margin upper clamp [K]
    DL_JKT_DB_LO    : REAL := 0.0;          // 死区域下限（Deadband lower clamp）[%] / Deadband lower clamp [%]
    DL_JKT_DB_HI    : REAL := 10.0;                // 死区域上限（Deadband upper clamp）[%] / Deadband upper clamp [%]
    DL_JKT_HYST     : REAL := 0.5;          // 触限回差（Limit hysteresis）[K]，防边界抖动 / Limit hysteresis [K]
    DL_JKT_K_PER_PCT : REAL := 0.5;         // 阀位传热增益（K per percent）[K/%]，偏离留档③ / Heat gain per percent [K/%]
    DL_JKT_MIN_PER_H : REAL := 60.0;        // 分钟换算（Minutes per hour）[-] / Minutes per hour
    DL_JKT_MS_PER_MIN : REAL := 60000.0;    // 毫秒→分钟换算（Milliseconds-to-minutes scale）[-] / Milliseconds-to-minutes scale
    DL_JKT_OPEN_EPS : REAL := 0.5;          // 「阀已开」判据（Valve open epsilon）[%] / Valve open epsilon [%]
    DL_JKT_ERR_NONFIN : UDINT := 16#0005_02FC; // 0005_02FC 温度或 PID 输出非有限【故障级】/ Non-finite temperature or PID output
    DL_JKT_ERR_REV    : UDINT := 16#0005_02FD; // 0005_02FD 温差为负且要求升温（传感器反装）【故障级】/ Reversed sensor, fault level
    DL_JKT_ERR_STATE  : UDINT := 16#0005_02FE; // 0005_02FE 非法状态兜底【故障级】/ Illegal state fallback, fault level
    DL_JKT_INFO_LIM   : UDINT := 16#0005_01CF; // 0005_01CF 温差达上限升温侧冻结【信息级】/ Delta-T limit reached, info level
    DL_JKT_INFO_OT    : UDINT := 16#0005_01D0; // 0005_01D0 釜温超设定加裕量强制冷却【信息级】/ Over temperature, info level
    DL_JKT_INFO_SPLIT : UDINT := 16#0005_01D1; // 0005_01D1 分程重叠区被死区分离【信息级】/ Split-range overlap separated, info level
END_VAR

// ============================================================================
// 段 1｜实例无条件周期刷新（R7/0.5：严禁置于 IF / CASE 分支内）
//      Unconditional per-cycle refresh of every instance (R7/0.5)
// ============================================================================
_fbTrigReset(CLK := bReset);                    // 复位上升沿（Reset rising edge）
_bResetEdge := _fbTrigReset.Q;                  // 复位单拍标志紧随实例赋值（R25 自清点）
_fbTonRate(
    IN := (NOT _bRateBreak),                    // 断输入拍串入 IN（R40 合规指纹）/ Window break folded into IN
    PT := tRateWindow
);                                              // 变化率统计窗（Rate window）

// 本拍码与条件预置（每拍重算；故障码以上拍锁存续用）
// Per-scan preset of codes and conditions, the fault code is carried from the latch
_uFaultCode := _uFaultLatched;                  // 故障码续用（Carry the latched fault code）
_uInfoCode  := 16#0000_0000;                    // 信息级码预清零（Info code preset to zero）
_bFaultCond := FALSE;                           // 故障条件预清零（Fault condition preset FALSE）
_fHeatTgt   := 0.0;                             // 热路目标预置 0（Heat target preset to zero）
_fCoolTgt   := 0.0;                             // 冷路目标预置 0（Cool target preset to zero）
_bLimitActive := FALSE;                         // 约束路径预置假（Limiting path preset FALSE）

// ============================================================================
// 段 2｜复位通道（R39：置于 CASE 之前，且不被掉使能分支屏蔽）
//      Reset path, before CASE and never masked by the disable branch
// ============================================================================
IF _bRateBreak THEN
    _bRateBreak := FALSE;                       // 统计窗断输入拍自清（Window break self-cleared）
END_IF

IF _bResetEdge THEN
    _bLimitLatched    := FALSE;                 // 触限锁存清除（Limit latch cleared）
    _bOverTempLatched := FALSE;                 // 超温锁存清除（Over-temp latch cleared）
    _fRateMeasInt     := 0.0;                   // 变化率测量值清零（Rate measurement cleared）
    _fDtWinStart      := 0.0;                   // 窗起点清零（Window start cleared）
    _bRateInit        := FALSE;                 // 窗首扫标志复位，重装基准（Init flag reset, R41）
    _uFaultLatched    := 16#0000_0000;          // 故障码锁存清除（Latched fault code cleared）
    _uFaultCode       := 16#0000_0000;          // 本拍故障码清空，防止段6 重新锁存旧码（Clear this scan code）
    IF _eState = E_DL_JacketState.eFault THEN
        _eState := E_DL_JacketState.eIdle;      // 故障态回空闲（Fault state back to idle）
        _bFaultCond := FALSE;                   // 故障条件清除（Fault condition cleared）
    END_IF
END_IF

// ============================================================================
// 段 3｜输入防御与参数钳位（镜像量每拍只锁一次，R38）
//      Input defense and parameter clamping, each mirror value latched once (R38)
// ============================================================================
IF (NOT (fReactorTemp >= DL_JKT_TEMP_MIN AND fReactorTemp <= DL_JKT_TEMP_MAX))
OR (NOT (fJacketTemp >= DL_JKT_TEMP_MIN AND fJacketTemp <= DL_JKT_TEMP_MAX))
OR (NOT (fPidOut >= (-DL_JKT_PID_MAX) AND fPidOut <= DL_JKT_PID_MAX)) THEN
    _bFaultCond := TRUE;                        // 非有限或越域即故障（Non-finite or out-of-domain is a fault）
    _uFaultCode := DL_JKT_ERR_NONFIN;           // 0005_02FC 温度或 PID 输出非有限【故障级】/ Non-finite input, fault level
    _fReactorNow := 0.0;                        // 快照置零，绝不用脏值（Snapshots zeroed）
    _fJacketNow  := 0.0;                        // 夹套快照置零（Jacket snapshot zeroed）
    _fPidNow     := 0.0;                        // PID 快照置零（PID snapshot zeroed）
ELSE
    _fReactorNow := fReactorTemp;               // 釜温快照（Reactor snapshot）
    _fJacketNow  := fJacketTemp;                // 夹套温快照（Jacket snapshot）
    _fPidNow     := fPidOut;                    // PID 快照（PID snapshot）
END_IF

// 参数域钳位（R35：守卫、封顶与判据同向）
// Parameter clamping so that guard, ceiling and comparison stay in step (R35)
_fDeltaTMaxEff := LIMIT(DL_JKT_DT_LO, fDeltaTMax, DL_JKT_DT_HI);        // 温差上限 5~150 K（Delta-T limit clamped）
_fRateLimEff   := LIMIT(DL_JKT_RATE_LO, fDeltaTRate, DL_JKT_RATE_HI);   // 变化率 0.1~50 K/min（Rate limit clamped）
_fOtMarginEff  := LIMIT(DL_JKT_OT_LO, fOverTempMargin, DL_JKT_OT_HI);   // 超温裕量 0.5~50 K（Margin clamped）
_fDeadbandEff  := LIMIT(DL_JKT_DB_LO, fDeadband, DL_JKT_DB_HI);         // 死区 0~10 %（Deadband clamped）
_fOutLowEff    := fOutMin;                      // 输出下限取引脚值（Output low taken from the pin）
_fOutHighEff   := fOutMax;                      // 输出上限取引脚值（Output high taken from the pin）
IF _fOutLowEff > _fOutHighEff THEN
    _fSwapTmp    := _fOutLowEff;                // 交换临时量（Swap scratch）
    _fOutLowEff  := _fOutHighEff;               // 下限取原上限（Low takes the former high）
    _fOutHighEff := _fSwapTmp;                  // 上限取原下限（High takes the former low）
END_IF

// 温差→阀位速率折算（偏离留档③）：[%/s] = (K/min ÷ 60) ÷ (K/%)
// Delta-T rate converted into an output rate in percent per second
IF _fRateLimEff > DL_JKT_EPS THEN
    _fRatePctS := (_fRateLimEff / DL_JKT_MIN_PER_H) / DL_JKT_K_PER_PCT;  // 折算（Converted rate）
ELSE
    _fRatePctS := 0.0;                          // 非法值按 0（限速器把 0 视为不限，防御性兜底）
END_IF

// ============================================================================
// 段 4｜温差与变化率测量（窗内斜率；窗边界断输入一拍，R40/R42）
//      Delta-T and its rate; the window boundary breaks the timer input for one scan
// ============================================================================
fDeltaT := _fReactorNow - _fJacketNow;          // 温差 = 釜温 − 夹套温（Delta-T, signed）
_fRateMin := TIME_TO_REAL(tRateWindow) / DL_JKT_MS_PER_MIN;  // 窗口分钟值（Window in minutes）
IF NOT _bRateInit THEN
    _bRateInit   := TRUE;                       // 首扫只装基准（R19：只装基准，不做判据）
    _fDtWinStart := fDeltaT;                    // 窗起点取首拍温差（Seed the window with the first scan value）
END_IF
IF _fbTonRate.Q THEN
    IF _fRateMin > DL_JKT_EPS THEN
        _fRateMeasInt := (fDeltaT - _fDtWinStart) / _fRateMin;  // 窗内平均斜率（Mean slope in the window）
    ELSE
        _fRateMeasInt := 0.0;                   // 窗长非法不出率（Illegal window, no rate）
    END_IF
    _fDtWinStart := fDeltaT;                    // 新窗起点（New window start）
    _bRateBreak  := TRUE;                       // 断输入一拍，ET 归零（R40）
END_IF

// ============================================================================
// 段 5｜状态机（约束层 + 分程层；ENUM + CASE，含 ELSE 兜底）
//      State machine: constraint layer plus split-range layer
// ============================================================================
// 5.1 温差触限与超温判定（回差防边界抖动）
//     Delta-T limit and over-temperature with hysteresis
IF fDeltaT >= _fDeltaTMaxEff THEN
    _bLimitLatched := TRUE;                     // 达上限即锁存（Reach the limit, latch it）
ELSIF fDeltaT < (_fDeltaTMaxEff - DL_JKT_HYST) THEN
    _bLimitLatched := FALSE;                    // 回落超回差才解除（Release only beyond the hysteresis）
END_IF
IF _fReactorNow > (fTempSetpoint + _fOtMarginEff) THEN
    _bOverTempLatched := TRUE;                  // 超温锁存（Over temperature latched）
    _uInfoCode := DL_JKT_INFO_OT;               // 0005_01D0 超温强制冷却【信息级】/ Over temperature
ELSIF _fReactorNow < (fTempSetpoint + _fOtMarginEff - DL_JKT_HYST) THEN
    _bOverTempLatched := FALSE;                 // 回落超回差才解除（Release only beyond the hysteresis）
END_IF

// 5.2 反装判据：温差为负且要求升温（本件最有价值的一条）
//     Reversed-sensor criterion: negative delta-T while heating is demanded
IF (NOT _bFaultCond) AND (fDeltaT < (-DL_JKT_HYST)) AND (_fPidNow > _fDeadbandEff) THEN
    _bFaultCond := TRUE;                        // 传感器疑似反装（Sensor likely reversed）
    _uFaultCode := DL_JKT_ERR_REV;              // 0005_02FD 温差为负且要求升温【故障级】/ Reversed sensor, fault level
END_IF

// 5.3 约束路径标记：触限、超温，或限速器仍在追赶（保证退出约束时平滑回收，不回跳）
//     Limiting path flag: limit active, over temperature, or the limiter still catching up
_bLimitActive := _bLimitLatched OR _bOverTempLatched
              OR _fbRlHeat.bLimiting OR _fbRlCool.bLimiting;

IF _bFaultCond THEN
    _eState := E_DL_JacketState.eFault;         // 故障条件优先于状态机（Fault outranks the machine）
END_IF

// 掉使能冻结分支：显式排除故障态（R39 合法写法①），复位通道仍可从故障态退出
// Disable branch explicitly excludes the fault state so the reset path still works
IF (NOT bEnable) AND (_eState <> E_DL_JacketState.eFault) THEN
    _eState := E_DL_JacketState.eIdle;          // 冻结回空闲（Freeze back to idle）
END_IF

CASE _eState OF

    E_DL_JacketState.eIdle: // 空闲：等使能与参数闸门
        IF bEnable AND (NOT _bFaultCond) THEN
            _eState := E_DL_JacketState.eHold;  // 进保持态等 PID 有效（Enter hold until the PID is valid）
        END_IF

    E_DL_JacketState.eHold: // 保持：两路 0，按 PID 与死区决定进入哪个方向
        _fHeatTgt := 0.0;                       // 热路目标 0（Heat target zero）
        _fCoolTgt := 0.0;                       // 冷路目标 0（Cool target zero）
        IF _bOverTempLatched THEN
            _eState   := E_DL_JacketState.eCool;    // 超温强制冷却（Forced cooling）
            _fCoolTgt := _fOutHighEff;          // 冷路给满量程（Cool at the upper limit）
        ELSIF _bLimitLatched THEN
            _eState := E_DL_JacketState.eHold;  // 触限期间保持冻结（Stay frozen while limited）
        ELSIF _fPidNow > _fDeadbandEff THEN
            _eState := E_DL_JacketState.eHeat;  // 要求升温（Heating demanded）
        ELSIF _fPidNow < (-_fDeadbandEff) THEN
            _eState := E_DL_JacketState.eCool;  // 要求冷却（Cooling demanded）
        ELSE
            _eState := E_DL_JacketState.eHold;  // 死区内保持（Inside the deadband)
        END_IF

    E_DL_JacketState.eHeat: // 升温：热路跟 PID，冷路 0
        _fCoolTgt := 0.0;                       // 冷路恒 0（Cool path forced zero）
        IF _bLimitLatched THEN
            _fHeatTgt := 0.0;                   // 触限冻结：目标 0，由限速器斜坡回落（Freeze, ramp down by the limiter）
            _uInfoCode := DL_JKT_INFO_LIM;      // 0005_01CF 温差达上限升温侧冻结【信息级】/ Delta-T limit reached
            _eState   := E_DL_JacketState.eHold;    // 进保持（Enter hold）
        ELSIF _bOverTempLatched THEN
            _fHeatTgt := 0.0;                   // 超温：热路目标 0（Over temperature, heat target zero）
            _eState   := E_DL_JacketState.eCool;    // 强制冷却（Forced cooling）
        ELSIF ABS(_fPidNow) <= _fDeadbandEff THEN
            _fHeatTgt := 0.0;                   // 死区内：热路目标 0（Inside the deadband）
            _eState   := E_DL_JacketState.eHold;    // 回保持（Back to hold）
            _uInfoCode := DL_JKT_INFO_SPLIT;    // 0005_01D1 分程重叠区被死区分离【信息级】/ Split-range overlap separated
        ELSE
            _fHeatTgt := LIMIT(_fOutLowEff, _fPidNow, _fOutHighEff);    // 热路跟 PID 并限幅（Heat follows the PID, clamped）
        END_IF

    E_DL_JacketState.eCool: // 冷却：冷路跟反相 PID，热路 0
        _fHeatTgt := 0.0;                       // 热路恒 0（Heat path forced zero）
        IF _bOverTempLatched THEN
            _fCoolTgt := _fOutHighEff;          // 超温：冷路给满（Cool at the upper limit）
            _uInfoCode := DL_JKT_INFO_OT;       // 0005_01D0 超温强制冷却【信息级】/ Over temperature
        ELSIF _fReactorNow < fTempSetpoint THEN
            _fCoolTgt := 0.0;                   // 釜温低于设定：停冷（Below setpoint, cooling stops）
            _eState   := E_DL_JacketState.eHold;    // 回保持（Back to hold）
        ELSIF ABS(_fPidNow) <= _fDeadbandEff THEN
            _fCoolTgt := 0.0;                   // 死区内：冷路目标 0（Inside the deadband）
            _eState   := E_DL_JacketState.eHold;    // 回保持（Back to hold）
            _uInfoCode := DL_JKT_INFO_SPLIT;    // 0005_01D1 分程重叠区被死区分离【信息级】/ Split-range overlap separated
        ELSE
            _fCoolTgt := LIMIT(_fOutLowEff, 0.0 - _fPidNow, _fOutHighEff);  // 冷路取反相 PID 并限幅（Cool takes the inverted PID, clamped）
        END_IF

    E_DL_JacketState.eFault: // 故障：两路强制 0，等复位沿（段2）
        _fHeatTgt := 0.0;                       // 热路目标 0（Heat target zero）
        _fCoolTgt := 0.0;                       // 冷路目标 0（Cool target zero）

    ELSE // 兜底：非法状态
        _uFaultCode := DL_JKT_ERR_STATE;        // 0005_02FE 非法状态兜底【故障级】/ Illegal state fallback
        _bFaultCond := TRUE;                    // 置故障条件（Raise the fault condition）
        _eState     := E_DL_JacketState.eFault; // 强制回故障态（Force the fault state）
        _fHeatTgt   := 0.0;                     // 热路目标 0（Heat target zero）
        _fCoolTgt   := 0.0;                     // 冷路目标 0（Cool target zero）
END_CASE

// ============================================================================
// 段 6｜冷热分程限速（组合调用 FB_DL_RateLimiter，算法在低层件内，绝不内联）
//      Split-range rate limiting by composing the low-level limiter, never inlined
//      未受限时 bTrack = TRUE（输出等于输入，无扰直通）；受限时 bTrack = FALSE，
//      按 _fRatePctS（由 fDeltaTRate 折算）限速，退出跟踪那一拍从当前值开始，不回跳。
//      Unconstrained passes through, constrained ramps from the present value
// ============================================================================
_fbRlHeat(
    bEnable     := TRUE,
    fIn         := _fHeatTgt,
    fRateUp     := _fRatePctS,
    fRateDown   := _fRatePctS,
    bTrack      := (NOT _bLimitActive) OR (NOT bEnable),
    fTrackValue := _fHeatTgt,
    tSampleTime := tCycle
);                                              // 热路限速（Heat path rate limiting）
_fbRlCool(
    bEnable     := TRUE,
    fIn         := _fCoolTgt,
    fRateUp     := _fRatePctS,
    fRateDown   := _fRatePctS,
    bTrack      := (NOT _bLimitActive) OR (NOT bEnable),
    fTrackValue := _fCoolTgt,
    tSampleTime := tCycle
);                                              // 冷路限速（Cool path rate limiting）

// ============================================================================
// 段 7｜码位单一优先级链（全拍只写一次，信息级不置 bError）
//      Single priority chain for the codes, written once per scan
// ============================================================================
IF _uFaultCode <> 16#0000_0000 THEN
    _uFaultLatched := _uFaultCode;              // 故障码锁存（Latched until reset）
    uErrorId  := _uFaultCode;                   // 故障级码优先（Fault-level code wins）
    uDiagCode := _uFaultCode;                   // 诊断码同源（Diagnostic code mirrors the fault）
    bError    := TRUE;                          // 故障标志置位（Error flag raised）
ELSIF _uInfoCode <> 16#0000_0000 THEN
    uErrorId  := 16#0000_0000;                  // 信息级不占故障码（Info level leaves the fault code empty）
    uDiagCode := _uInfoCode;                    // 诊断码取信息级码（Diagnostic code takes the info code）
    bError    := FALSE;                         // 信息级不置故障位（Info level never raises the error flag）
ELSE
    uErrorId  := 16#0000_0000;                  // 无码（No code）
    uDiagCode := 16#0000_0000;                  // 无码（No code）
    bError    := FALSE;                         // 无故障（No error）
END_IF

// ============================================================================
// 段 8｜出口钳位与保持语义重写（R27/R43：结论逐拍重写，冷热互斥）
//      Output clamping and held-semantics rewrite, heat and cool mutually exclusive
// ============================================================================
_fHeatPrev := LIMIT(_fOutLowEff, _fbRlHeat.fOut, _fOutHighEff);     // 热路取限速器输出并夹域（Heat from the limiter, clamped）
_fCoolPrev := LIMIT(_fOutLowEff, _fbRlCool.fOut, _fOutHighEff);     // 冷路取限速器输出并夹域（Cool from the limiter, clamped）

// 互斥出口：决不允许冷热同开（同拍只保留一路，且优先保冷——冷却属安全方向）
// Mutual exclusion: heat and cool can never be open together, cooling wins as the safe direction
IF (_fHeatPrev > DL_JKT_OPEN_EPS) AND (_fCoolPrev > DL_JKT_OPEN_EPS) THEN
    _fHeatPrev := 0.0;                          // 两路同开：热路强制归零（Both open: heat forced to zero）
END_IF

fHeatOut      := _fHeatPrev;                    // 热路出口逐拍重写（Heat output rewritten every scan）
fCoolOut      := _fCoolPrev;                    // 冷路出口逐拍重写（Cool output rewritten every scan）
fDeltaTRateMeas := _fRateMeasInt;               // 变化率出口逐拍重写（Measured rate rewritten）
bDeltaTLimited := _bLimitLatched;               // 触限位逐拍重写（Limit flag rewritten）
bOverTemp     := _bOverTempLatched;             // 超温位逐拍重写（Over-temperature flag rewritten）
eVerdict      := _eState;                       // 执行方向逐拍重写（Verdict rewritten every scan）

// 健康态仲裁（引用属主 A1 的四态语言）
// Health arbitration mapped onto the A1 health language
IF _eState = E_DL_JacketState.eFault THEN
    eHealth := E_DL_Ne107Status.eFailure;       // 故障：温度或 PID 不可信（Failure）
ELSIF NOT bEnable THEN
    eHealth := E_DL_Ne107Status.eUnknown;       // 未知：未使能（Unknown）
ELSIF _bOverTempLatched THEN
    eHealth := E_DL_Ne107Status.eOutOfSpec;     // 越规：釜温越界（Out of spec）
ELSIF _bLimitLatched THEN
    eHealth := E_DL_Ne107Status.eMaintenanceReq;    // 需维护：温差约束长期生效，传热面可能结垢（Maintenance required）
ELSE
    eHealth := E_DL_Ne107Status.eOk;            // 正常（OK）
END_IF

END_FUNCTION_BLOCK
